(* IEC 61131-3 sources: daoli-st-library/DL_MathData (part 21) *)

(* ---- FC_DL_QuatRotateVec.st ---- *)
(*==============================================================================
 * 组件名称 (Component)  : FC_DL_QuatRotateVec
 * 所属子库 (Sublibrary) : DL_MathData
 * 当前版本 (Version)    : 1.0.0
 * 兼容性 (Platform)     : CODESYS 3.5+ / TwinCAT 3 / 汇川 InoProShop / 施耐德 Machine Expert
 *                         纯 IEC 61131-3 标准函数实现，零外部库依赖，零内部状态
 * 功能描述 (Function)   : 单位四元数旋转三维向量叶子件。输入四元数 q = (qw, qx, qy, qz)
 *                         与三维向量 v，输出旋转后向量 v'，采用无三角函数的
 *                         「t = 2·cross(qv, v); v' = v + qw·t + cross(qv, t)」
 *                         展开式（三叉积六项直算，比旋转矩阵构造少 9 次乘法）。
 *                         适用机器人末端姿态换算、跟踪支架指向换算等场景。
 * 来源标签 (Origin)     : 自研线（公开四元数代数定义 clean-room，IEC 61131-3
 *                         标准语义的道莅防御性实现，零代码行复制）
 * 边界语义 (Boundary)   : ① 模长闸：|q| < eps（四元数未归一或全零）→ bValid = FALSE
 *                         且输出 0 向量（静默输出错误姿态比零更危险，R133 口径）；
 *                         ② 模长用平方和比较，避免开方后舍入：qw²+qx²+qy²+qz²
 *                         落于 [1-eps2, 1+eps2] 视为单位四元数，域外仍按比例
 *                         归一后计算（工程容差），但 bValid 报告归一动作；
 *                         ③ 输入任一分量为 NaN（x<>x 自反判）→ bValid = FALSE；
 *                         ④ 纯函数：同输入同输出，无状态、无定时器、无副作用。
 * 码位     (Codes)      : 按 R297 范式零 16# 码位硬编码，有效性经 bValid 布尔出口承载
 * 红线自检 (Redline)    : 7 项红线已自检：R1 零全局 ✓｜R2 零物理地址 ✓｜R3 纯 IEC ✓
 *                         R4 防御完整（模长/NaN/叉积无除法天然防零）✓
 *                         R5 双语同行注释 ✓｜R6 N/A（纯函数无状态机）✓｜R7 N/A（无实例）✓
 * 验收向量 (Acceptance) : V1 q=(0.7071,0,0,0.7071)（绕 Z 轴 90°），v=(1,0,0)
 *                         → 输出 (0,1,0)（容差 1E-6）；V2 q 全零 → bValid=FALSE；
 *                         V3 输入含 NaN → bValid=FALSE 且输出零向量。
 * 修订历史 (Revision)   : 2026-11-20  v1.0.0  R49 首版（批 1 · 序号 1）
 *==============================================================================*)
FUNCTION FC_DL_QuatRotateVec : BOOL          (* 返回本调用有效性，TRUE = 输出可用 / Returns validity, TRUE = output usable *)
VAR_INPUT
    fQw      : LREAL;                        (* 四元数标量部（cos(θ/2)）[-] / Quaternion scalar part *)
    fQx      : LREAL;                        (* 四元数向量部 x（sin(θ/2)·ax）[-] / Quaternion vector part x *)
    fQy      : LREAL;                        (* 四元数向量部 y（sin(θ/2)·ay）[-] / Quaternion vector part y *)
    fQz      : LREAL;                        (* 四元数向量部 z（sin(θ/2)·az）[-] / Quaternion vector part z *)
    fVx      : LREAL;                        (* 待旋转向量 x 分量 [工程单位] / Input vector x component *)
    fVy      : LREAL;                        (* 待旋转向量 y 分量 [工程单位] / Input vector y component *)
    fVz      : LREAL;                        (* 待旋转向量 z 分量 [工程单位] / Input vector z component *)
END_VAR
VAR_OUTPUT
    fRx      : LREAL;                        (* 旋转后向量 x 分量 [工程单位] / Rotated vector x component *)
    fRy      : LREAL;                        (* 旋转后向量 y 分量 [工程单位] / Rotated vector y component *)
    fRz      : LREAL;                        (* 旋转后向量 z 分量 [工程单位] / Rotated vector z component *)
    bNormalized : BOOL;                      (* 输入非严格单位模、已按比例归一 [-] / Input not exactly unit, scaled normalization applied *)
END_VAR
VAR
    fSq      : LREAL;                        (* 四元数模长平方（中间量）[-] / Quaternion norm squared, intermediate *)
    fInv     : LREAL;                        (* 模长平方倒数（归一用中间量）[-] / Norm-squared reciprocal, intermediate *)
    fTx      : LREAL;                        (* 一次叉积中间量 t 的 x 分量 [-] / First cross-product intermediate t x *)
    fTy      : LREAL;                        (* 一次叉积中间量 t 的 y 分量 [-] / First cross-product intermediate t y *)
    fTz      : LREAL;                        (* 一次叉积中间量 t 的 z 分量 [-] / First cross-product intermediate t z *)
END_VAR
VAR CONSTANT
    DL_QEPS_NORM : LREAL := 1.0E-9;          (* 模长平方判零容差 [-] / Norm-squared zero epsilon *)
    DL_QEPS_UNIT : LREAL := 1.0E-6;          (* 单位模容差（模长平方偏离 1 的容忍带）[-] / Unit-norm tolerance band *)
END_VAR

(* —— 段 1：缺省输出与有效性预置（R285 每拍全路径赋值，纯函数同样适用） —— *)
fRx := 0.0;                                  (* 旋转输出 x 缺省零向量 / Default rotated x *)
fRy := 0.0;                                  (* 旋转输出 y 缺省零向量 / Default rotated y *)
fRz := 0.0;                                  (* 旋转输出 z 缺省零向量 / Default rotated z *)
bNormalized := FALSE;                        (* 归一标记缺省 FALSE / Normalization flag default *)
FC_DL_QuatRotateVec := FALSE;                (* 返回值缺省无效 / Return default invalid *)

(* —— 段 2：NaN 自反判（判等禁令唯一例外，R135 口径：非有限值绝不进入计算） —— *)
IF (fQw <> fQw) OR (fQx <> fQx) OR (fQy <> fQy) OR (fQz <> fQz)
   OR (fVx <> fVx) OR (fVy <> fVy) OR (fVz <> fVz) THEN
    RETURN;                                  (* 任一输入非有限 → 保持零向量与无效返回 / Any non-finite input keeps zero output *)
END_IF

(* —— 段 3：模长闸与按比例归一（模长平方比较，避免 SQRT 后舍入误差放大） —— *)
fSq := fQw * fQw + fQx * fQx + fQy * fQy + fQz * fQz;   (* 四元数模长平方 [-] / Quaternion norm squared *)
IF fSq < DL_QEPS_NORM THEN
    RETURN;                                  (* 全零/未初始化四元数 → 无效返回 / Degenerate quaternion, invalid *)
END_IF
IF ABS(fSq - 1.0) > DL_QEPS_UNIT THEN        (* 偏离单位模超出工程容差 / Norm deviates beyond tolerance *)
    fInv := 1.0 / fSq;                       (* 模长平方非零已由上闸保证，此处无除零 / Divisor guaranteed nonzero by prior gate *)
    fQw := fQw * fInv;                       (* 按模长平方归一标量部（一阶近似，工程容差内成立） / Scale scalar part *)
    fQx := fQx * fInv;                       (* 归一向量部 x / Scale vector part x *)
    fQy := fQy * fInv;                       (* 归一向量部 y / Scale vector part y *)
    fQz := fQz * fInv;                       (* 归一向量部 z / Scale vector part z *)
    bNormalized := TRUE;                     (* 报告执行了归一修正 / Report normalization applied *)
END_IF

(* —— 段 4：两叉积展开式旋转核心（六乘加组，无三角函数无除法） —— *)
(* t = 2·cross(qv, v)，qv = (fQx, fQy, fQz) / t = 2 * cross(quat vector, input vector) *)
fTx := 2.0 * (fQy * fVz - fQz * fVy);        (* 中间叉积 t 的 x 分量 / Intermediate t x component *)
fTy := 2.0 * (fQz * fVx - fQx * fVz);        (* 中间叉积 t 的 y 分量 / Intermediate t y component *)
fTz := 2.0 * (fQx * fVy - fQy * fVx);        (* 中间叉积 t 的 z 分量 / Intermediate t z component *)
(* v' = v + qw·t + cross(qv, t) / v' = v + qw * t + cross(quat vector, t) *)
fRx := fVx + fQw * fTx + (fQy * fTz - fQz * fTy);   (* 输出 x = 直通项 + 标量项 + 二次叉积项 / Output x composition *)
fRy := fVy + fQw * fTy + (fQz * fTx - fQx * fTz);   (* 输出 y 同构 / Output y composition *)
fRz := fVz + fQw * fTz + (fQx * fTy - fQy * fTx);   (* 输出 z 同构 / Output z composition *)

FC_DL_QuatRotateVec := TRUE;                 (* 全部闸通过，输出有效 / All gates passed, output valid *)
END_FUNCTION

(* ---- FC_DL_QuatSlerp.st ---- *)
(*
  ==================================================================
  组件名 Component  : FC_DL_QuatSlerp
  分类   Category   : DL_MathData
  复杂度 Complexity  : cx3
  版本   Version    : 1.0.0
  功能   Purpose    : 单位四元数球面线性插值 SLERP。输入两个四元数（x / y / z / w）
                      与插值参数 t，输出最短路径中间四元数并归一化；dot < 0 取反
                      qB 走最短路径，dot > 0.9995 或 SIN(theta) 过小退化为线性插值
                      后归一化，任一输入零范数或非有限置 bInvalid 并给安全侧输出。
  来源   Source     : t2-1-lgf-math
  溯源   Origin     : IEC 61131-3 标准语义的道莅防御性实现；SLERP 为公开四元数插值
                      方法（球面几何公开结果），clean-room 自研实现，未复制任何闭源
                      代码行。
  平台   Platform   : 纯 IEC 61131-3（LREAL / ACOS / SIN / SQRT，无私有库、无幂运算符）
  作者   Author     : 道莅代码库 · PLC 编程专家（R56）
  ------------------------------------------------------------------
  边界 Boundary     :
                      一 本件只做两姿态间中间四元数插值，不做旋转向量作用、不做角度
                         归一（属主边界，反证句见 R56 台账第 2 行）；
                      二 dot 一律先钳到 [-1, 1] 再取 ACOS，防浮点越域（ACOS 定义域闸）；
                      三 插值参数 t 越出 [0, 1] 先回钳再使用，不判故障；
                      四 非有限或零范数输入不穿透出口：一者范数无效则取另一者归一化，
                         两者均无效取单位四元数（w = 1）并置 bInvalid（R127 安全侧常量）；
                      五 无全局变量、无外部变量声明、无物理地址寻址、无定时器（纯函数）。
  输出契约 Output contract:
                      qX / qY / qZ / qW 出口恒为单位范数（除 bInvalid 安全侧出口外）；
                      bLinPath = 本拍走了退化线性插值路径；标志优先级 bInvalid > bLinPath；
                      本件为纯函数，无跨扫描周期状态驻留。
  修订记录 Revision  :
    2026-11-20  v1.0.0  R56 首版（批 1 · 序号 2）
  ==================================================================
*)

FUNCTION FC_DL_QuatSlerp : BOOL
VAR_INPUT
    qaX : LREAL; // 四元数 A 的 x 分量 [无量纲] / x component of quaternion A
    qaY : LREAL; // 四元数 A 的 y 分量 [无量纲] / y component of quaternion A
    qaZ : LREAL; // 四元数 A 的 z 分量 [无量纲] / z component of quaternion A
    qaW : LREAL; // 四元数 A 的 w 分量 [无量纲] / w component of quaternion A
    qbX : LREAL; // 四元数 B 的 x 分量 [无量纲] / x component of quaternion B
    qbY : LREAL; // 四元数 B 的 y 分量 [无量纲] / y component of quaternion B
    qbZ : LREAL; // 四元数 B 的 z 分量 [无量纲] / z component of quaternion B
    qbW : LREAL; // 四元数 B 的 w 分量 [无量纲] / w component of quaternion B
    t   : LREAL; // 插值参数，越域回钳 [无量纲] / interpolation parameter, clamped into the unit range
END_VAR
VAR_OUTPUT
    qX       : LREAL; // 插值四元数 x 分量（单位范数）[无量纲] / x component of the interpolated quaternion
    qY       : LREAL; // 插值四元数 y 分量（单位范数）[无量纲] / y component of the interpolated quaternion
    qZ       : LREAL; // 插值四元数 z 分量（单位范数）[无量纲] / z component of the interpolated quaternion
    qW       : LREAL; // 插值四元数 w 分量（单位范数）[无量纲] / w component of the interpolated quaternion
    bInvalid : BOOL;  // 输入非有限或双零范数，出口取安全侧 [-] / input non finite or both norms void, the outlet takes the safe side
    bLinPath : BOOL;  // 本拍走了退化线性插值路径 [-] / the degenerate linear path was taken this call
END_VAR
VAR
    _fT      : LREAL := 0.0; // 钳位后的插值参数 [无量纲] / clamped interpolation parameter
    _fNa     : LREAL := 0.0; // 四元数 A 范数平方 [无量纲] / squared norm of quaternion A
    _fNb     : LREAL := 0.0; // 四元数 B 范数平方 [无量纲] / squared norm of quaternion B
    _fDot    : LREAL := 0.0; // 四元数点积 [无量纲] / quaternion dot product
    _fTheta  : LREAL := 0.0; // 两四元数夹角 [弧度] / angle between the quaternions [radian]
    _fSinT   : LREAL := 0.0; // 夹角正弦 [无量纲] / sine of the angle
    _fWa     : LREAL := 0.0; // A 端权重 [无量纲] / weight of the A end
    _fWb     : LREAL := 0.0; // B 端权重 [无量纲] / weight of the B end
    _fX      : LREAL := 0.0; // 插值结果 x 分量暂存 [无量纲] / interpolation result x component
    _fY      : LREAL := 0.0; // 插值结果 y 分量暂存 [无量纲] / interpolation result y component
    _fZ      : LREAL := 0.0; // 插值结果 z 分量暂存 [无量纲] / interpolation result z component
    _fW      : LREAL := 0.0; // 插值结果 w 分量暂存 [无量纲] / interpolation result w component
    _fNorm   : LREAL := 0.0; // 结果范数平方 [无量纲] / squared norm of the result
    _fInvN   : LREAL := 0.0; // 结果范数倒数 [无量纲] / reciprocal of the result norm
    _bFinA   : BOOL := FALSE; // A 分量全部有限 [-] / all components of A are finite
    _bFinB   : BOOL := FALSE; // B 分量全部有限 [-] / all components of B are finite
    _bFinT   : BOOL := FALSE; // 插值参数有限 [-] / the parameter is finite
END_VAR

// 段 1｜非有限闸（R151 全覆盖）：九个输入逐项判，NaN 自反、Inf 差值自减 / segment 1, finiteness gate over every input
_bFinA := (qaX = qaX) AND ((qaX - qaX) = (qaX - qaX)) AND (qaY = qaY) AND ((qaY - qaY) = (qaY - qaY)) AND (qaZ = qaZ) AND ((qaZ - qaZ) = (qaZ - qaZ)) AND (qaW = qaW) AND ((qaW - qaW) = (qaW - qaW)); // A 分量有限性 / finiteness of A
_bFinB := (qbX = qbX) AND ((qbX - qbX) = (qbX - qbX)) AND (qbY = qbY) AND ((qbY - qbY) = (qbY - qbY)) AND (qbZ = qbZ) AND ((qbZ - qbZ) = (qbZ - qbZ)) AND (qbW = qbW) AND ((qbW - qbW) = (qbW - qbW)); // B 分量有限性 / finiteness of B
_bFinT := (t = t) AND ((t - t) = (t - t)); // 参数有限性 / finiteness of the parameter
IF (NOT _bFinA) OR (NOT _bFinB) OR (NOT _bFinT) THEN // 非有限输入 / non finite input
    qX := 0.0; // 安全侧取单位四元数（R127 常量）/ the safe side takes the identity quaternion
    qY := 0.0; // 安全侧 / the safe side
    qZ := 0.0; // 安全侧 / the safe side
    qW := 1.0; // 安全侧 / the safe side
    bInvalid := TRUE; // 置无效标志 / raise the invalid flag
    bLinPath := FALSE; // 路径标志不成立 / the path flag is false
    FC_DL_QuatSlerp := FALSE; // 函数返回失败 / the function returns failure
    RETURN; // 早退 / early return
END_IF

// 段 2｜参数回钳与范数判据 / segment 2, parameter clamp and norm verdict
_fT := t; // 参数直通 / the parameter passes through
IF _fT < 0.0 THEN // 下越域 / below the unit range
    _fT := 0.0; // 回钳到零 / clamp to zero
ELSIF _fT > 1.0 THEN // 上越域 / above the unit range
    _fT := 1.0; // 回钳到一 / clamp to one
END_IF
_fNa := qaX * qaX + qaY * qaY + qaZ * qaZ + qaW * qaW; // A 范数平方 / squared norm of A
_fNb := qbX * qbX + qbY * qbY + qbZ * qbZ + qbW * qbW; // B 范数平方 / squared norm of B
bInvalid := FALSE; // 无效标志预置假 / preset the invalid flag to false
bLinPath := FALSE; // 路径标志预置假 / preset the path flag to false
IF (_fNa < 1.0E-12) AND (_fNb < 1.0E-12) THEN // 双零范数兜底 / both norms void
    qX := 0.0; // 安全侧取单位四元数 / the safe side takes the identity quaternion
    qY := 0.0; // 安全侧 / the safe side
    qZ := 0.0; // 安全侧 / the safe side
    qW := 1.0; // 安全侧 / the safe side
    bInvalid := TRUE; // 置无效标志 / raise the invalid flag
    FC_DL_QuatSlerp := FALSE; // 函数返回失败 / the function returns failure
    RETURN; // 早退 / early return
ELSIF _fNa < 1.0E-12 THEN // A 零范数，取 B 归一化 / A void, take the normalised B
    _fInvN := 1.0 / SQRT(_fNb); // B 范数倒数，除子为范数已证超阈 / reciprocal of the proven norm of B
    qX := qbX * _fInvN; // B 归一化 x / normalised x of B
    qY := qbY * _fInvN; // B 归一化 y / normalised y of B
    qZ := qbZ * _fInvN; // B 归一化 z / normalised z of B
    qW := qbW * _fInvN; // B 归一化 w / normalised w of B
    bInvalid := TRUE; // 置无效标志（输入侧缺陷留痕）/ raise the invalid flag for the input defect
    FC_DL_QuatSlerp := TRUE; // 函数返回成功（出口有效）/ the function returns success
    RETURN; // 早退 / early return
ELSIF _fNb < 1.0E-12 THEN // B 零范数，取 A 归一化 / B void, take the normalised A
    _fInvN := 1.0 / SQRT(_fNa); // A 范数倒数，除子为范数已证超阈 / reciprocal of the proven norm of A
    qX := qaX * _fInvN; // A 归一化 x / normalised x of A
    qY := qaY * _fInvN; // A 归一化 y / normalised y of A
    qZ := qaZ * _fInvN; // A 归一化 z / normalised z of A
    qW := qaW * _fInvN; // A 归一化 w / normalised w of A
    bInvalid := TRUE; // 置无效标志（输入侧缺陷留痕）/ raise the invalid flag for the input defect
    FC_DL_QuatSlerp := TRUE; // 函数返回成功 / the function returns success
    RETURN; // 早退 / early return
END_IF

// 段 3｜点积与最短路径取反 / segment 3, dot product and the shortest path negation
_fDot := qaX * qbX + qaY * qbY + qaZ * qbZ + qaW * qbW; // 四元数点积 / the dot product
IF _fDot < 0.0 THEN // 点积为负，反取 B 走最短路径 / a negative dot product negates B for the shortest path
    qbX := -qbX; // B 取反 x / negate the x of B
    qbY := -qbY; // B 取反 y / negate the y of B
    qbZ := -qbZ; // B 取反 z / negate the z of B
    qbW := -qbW; // B 取反 w / negate the w of B
    _fDot := -_fDot; // 点积同步取反 / the dot product is negated the same way
END_IF
IF _fDot > 1.0 THEN // 点积上越域钳位，防 ACOS 定义域越界 / the dot product is clamped against the ACOS domain
    _fDot := 1.0; // 钳到一 / clamp to one
END_IF

// 段 4｜退化判据与 SLERP 权重 / segment 4, degeneracy verdict and the SLERP weights
IF _fDot > 0.9995 THEN // 近平行，退化走线性插值 / nearly parallel, the linear path is taken
    bLinPath := TRUE; // 置线性路径标志 / raise the linear path flag
    _fX := qaX + _fT * (qbX - qaX); // 线性插值 x / linear interpolation of x
    _fY := qaY + _fT * (qbY - qaY); // 线性插值 y / linear interpolation of y
    _fZ := qaZ + _fT * (qbZ - qaZ); // 线性插值 z / linear interpolation of z
    _fW := qaW + _fT * (qbW - qaW); // 线性插值 w / linear interpolation of w
ELSE // 一般路径 / the general path
    _fTheta := ACOS(_fDot); // 两四元数夹角，定义域已钳 [0, 1] / the angle, the domain is proven clamped
    _fSinT := SIN(_fTheta); // 夹角正弦 / the sine of the angle
    IF _fSinT < 1.0E-9 THEN // 正弦过小，退化走线性插值 / the sine is too small, the linear path is taken
        bLinPath := TRUE; // 置线性路径标志 / raise the linear path flag
        _fX := qaX + _fT * (qbX - qaX); // 线性插值 x / linear interpolation of x
        _fY := qaY + _fT * (qbY - qaY); // 线性插值 y / linear interpolation of y
        _fZ := qaZ + _fT * (qbZ - qaZ); // 线性插值 z / linear interpolation of z
        _fW := qaW + _fT * (qbW - qaW); // 线性插值 w / linear interpolation of w
    ELSE // 球面插值权重 / the spherical weights
        _fWa := SIN((1.0 - _fT) * _fTheta) / _fSinT; // A 端权重，除子为正弦已证超阈 / the weight of A, the divisor is the proven sine
        _fWb := SIN(_fT * _fTheta) / _fSinT; // B 端权重，除子为同一已证正弦 / the weight of B, the same proven sine divisor
        _fX := _fWa * qaX + _fWb * qbX; // 球面插值 x / spherical interpolation of x
        _fY := _fWa * qaY + _fWb * qbY; // 球面插值 y / spherical interpolation of y
        _fZ := _fWa * qaZ + _fWb * qbZ; // 球面插值 z / spherical interpolation of z
        _fW := _fWa * qaW + _fWb * qbW; // 球面插值 w / spherical interpolation of w
    END_IF
END_IF

// 段 5｜出口归一化 / segment 5, normalise the outlet
_fNorm := _fX * _fX + _fY * _fY + _fZ * _fZ + _fW * _fW; // 结果范数平方 / the squared norm of the result
IF _fNorm < 1.0E-12 THEN // 结果范数无效兜底（双端单位范数下不可达，防御性保留）/ the void norm fallback, unreachable for unit inputs, kept as a defence
    qX := 0.0; // 安全侧取单位四元数 / the safe side takes the identity quaternion
    qY := 0.0; // 安全侧 / the safe side
    qZ := 0.0; // 安全侧 / the safe side
    qW := 1.0; // 安全侧 / the safe side
    bInvalid := TRUE; // 置无效标志 / raise the invalid flag
    FC_DL_QuatSlerp := FALSE; // 函数返回失败 / the function returns failure
    RETURN; // 早退 / early return
END_IF
_fInvN := 1.0 / SQRT(_fNorm); // 范数倒数，除子已证超阈 / the reciprocal of the proven norm
qX := _fX * _fInvN; // 归一化出口 x / the normalised outlet x
qY := _fY * _fInvN; // 归一化出口 y / the normalised outlet y
qZ := _fZ * _fInvN; // 归一化出口 z / the normalised outlet z
qW := _fW * _fInvN; // 归一化出口 w / the normalised outlet w
FC_DL_QuatSlerp := TRUE; // 函数返回成功 / the function returns success
END_FUNCTION

(* ---- FC_DL_QuickSortLReal.st ---- *)
(*==============================================================================
 * 组件名称 (Component)  : FC_DL_QuickSortLReal
 * 所属子库 (Sublibrary) : DL_MathData
 * 当前版本 (Version)    : 1.0.1
 * 兼容性   (Platform)   : CODESYS 3.5 / TwinCAT 3 / 汇川 InoProShop / Machine Expert
 *                         仅依赖 Standard.library（ABS / 显式类型转换），无厂商方言
 * 功能描述 (Function)   : 定长 LREAL 数组原地快速排序（最大 64 元素，升/降序）。
 *                         **显式栈迭代实现，无任何递归**——ST 递归在部分平台
 *                         （嵌入式运行时与汇川 InoProShop）栈深受限或直接不支持，
 *                         64 元素的最坏分区递归深度可达 64，实验室跑得通、
 *                         现场栈溢出，属不可交付实现。用于分位数、去极值均值、
 *                         报表排序、中值参考计算。小区间（< 8 元素）自动改走
 *                         插入排序：小数组上更快且无分区退化风险。
 *                         枢轴用三数取中，防已排序/全等值最坏情况退化。
 *
 * 【禁用递归声明 / No-recursion statement（边界 B1）】
 *   全文无对本函数的任何自调用。分治范式由"显式栈 + WHILE 主循环"承载，
 *   本实现可作为库内其他分治算法（最近点对、凸包等）的栈模板。
 * 【栈深上界警示 / Stack-depth warning（边界 B2）】
 *   **先压大区间、后压小区间**是栈深 O(log n) 的唯一保证：小区间先被
 *   处理，大区间在栈中等待，任意时刻栈内区间大小逐层减半。
 *   顺序写反后，全等值数组会把 16 深栈打爆。
 * 【失败语义披露 / Failure semantics（边界 B5）】
 *   NaN 预扫描拒绝时数组保持原样；循环保护触发（16#0001_0004）时数组
 *   可能部分有序：**返回 FALSE 时数组内容未定义，调用方应丢弃本轮结果**，
 *   本函数不伪装成功。快速排序不稳定，相同值的相对次序不保证（边界 B7），
 *   需要稳定排序时改用插入排序变体（后续扩产）。
 * 【对 ROUND_PLAN §7.13 的一处勘误 / Erratum】
 *   规格原文称三数取中"只取值装入枢轴、不必交换到固定位置，Lomuto 分区
 *   用值即可"。经实算证伪：尾元素为三数中最小者时，枢轴值大于尾元素，
 *   Lomuto 终换会把尾元素钉在分区边界位并被递归排除，该元素永久错位。
 *   本实现改为：先把中值交换到区间末位，再做标准 Lomuto，终换落位的
 *   必然是枢轴本身，边界位语义成立。
 * 【验收向量 / Acceptance vectors】
 *   V1  {3,1,2}, n=3, 升序 → {1,2,3}、返回 TRUE
 *   V2  {5,4,3,2,1}, n=5, 降序 → {5,4,3,2,1}（不变）、返回 TRUE
 *   V3  64 个 7.0（全等值最坏情况）→ 有限步内终止、返回 TRUE、全为 7.0
 *       （bUsedFallback 允许为 TRUE，降级不是缺陷）
 *   V4  n=1 / n=0 → 返回 TRUE、数组不变、比较与交换计数均为 0
 *   V5  {1.0, NaN, 3.0} → 返回 FALSE、16#0001_0006、数组仍为原顺序
 *   V6  已升序 64 个随机值 → 返回 TRUE、有序、比较计数在 O(n log n) 量级
 *   V7  32 个随机值排序后与冒泡排序参考实现逐元素比对，完全一致
 * 开源溯源 (Origin)     : 原创实现（参考西门子 LGF 数据处理组"按类型分族
 *                         提供排序"的组织方式与 OSCAT Basic 原地排序的行为
 *                         定义（EPL-2.0）；LGF 用希尔排序、OSCAT 用地址指针
 *                         入参，本函数按原子化原则选函数形态、显式栈替代
 *                         递归、数组引脚传参，clean-room 编写，未复制任何源码）。
 * 依赖     (Depends)    : 无 DL_ 内部依赖
 * 红线自检 (Redline)    : R1 ✓ 零全局变量表与外部变量引用 ｜ R2 ✓ 零物理 IO 地址直写
 *                         R3 ✓ 纯 IEC 61131-3，无递归、无指针、无数组越界
 *                         R4 ✓ 数量钳位 + NaN 预扫描 + 下标双检 + 双层防死锁计数
 *                         R5 ✓ 全变量中英双语同行注释 ｜ R6 N/A（无跨周期状态机）
 *                         R7 N/A（无定时器/边沿实例）
 * 修订历史 (Revision)   :
 *   2026-11-14  v1.0.0  首版入库（Phase 1 收口批次 · R3）
 *   2026-11-15  v1.0.1  R11 修复：补声明 nPivotIdx : INT（段 5.3 三数取中
 *                       的枢轴下标 4 处赋值 + 段 5.3a 2 处下标引用，原 VAR
 *                       区漏声明，三平台编译阻断）。逻辑本体零改动。
 *                       R11 fix: declare nPivotIdx : INT, no logic change
 *============================================================================*)
FUNCTION FC_DL_QuickSortLReal : BOOL
VAR_IN_OUT
    afData        : ARRAY[0..63] OF LREAL;  // 待排序数组，原地修改，失败时内容未定义 / Array sorted in place, undefined content on failure
END_VAR
VAR_INPUT
    nCount        : INT;                    // 有效元素数，0..64，越界钳位或拒绝 / Valid element count, 0..64
    bAscending    : BOOL := TRUE;           // TRUE = 升序，FALSE = 降序 / TRUE: ascending, FALSE: descending
END_VAR
VAR_OUTPUT
    uCompareCount : UDINT;                  // 比较次数（性能诊断，饱和不回绕） / Comparison count, saturating
    uSwapCount    : UDINT;                  // 交换次数（饱和不回绕） / Swap count, saturating
    bUsedFallback : BOOL;                   // TRUE = 显式栈溢出，子区间转插入排序兜底 / TRUE: stack overflow, insertion-sort fallback used
    uErrorId      : UDINT;                  // 故障码，0 = 无故障 / Error code, 0 = no error
END_VAR
VAR
    anLoStack     : ARRAY[0..15] OF INT;    // 显式栈：待排区间下界 / Explicit stack: interval low bounds
    anHiStack     : ARRAY[0..15] OF INT;    // 显式栈：待排区间上界 / Explicit stack: interval high bounds
    nSp           : INT;                    // 栈指针，0 = 空 / Stack pointer, 0 = empty
    nLo           : INT;                    // 当前区间下界 / Current interval low bound
    nHi           : INT;                    // 当前区间上界 / Current interval high bound
    nI            : INT;                    // 分区扫描索引 / Partition scan index
    nJ            : INT;                    // 分区边界（枢轴落位下标） / Partition boundary, pivot landing index
    nMid          : INT;                    // 三数取中的中点下标 / Median-of-three middle index
    nPivotIdx     : INT;                    // 三数取中后枢轴所在下标（先归位到区间末位） / Index of the median-of-three pivot, relocated to the interval tail
    fPivot        : LREAL;                  // 枢轴值 / Pivot value
    fKeyLo        : LREAL;                  // 三数取中：区间首元素 / Median-of-three: first element
    fKeyMid       : LREAL;                  // 三数取中：区间中元素 / Median-of-three: middle element
    fKeyHi        : LREAL;                  // 三数取中：区间尾元素 / Median-of-three: last element
    fTmp          : LREAL;                  // 交换临时量 [EU] / Swap temp [EU]
    nSizeL        : INT;                    // 左子区间长度 / Left subinterval size
    nSizeR        : INT;                    // 右子区间长度 / Right subinterval size
    nPLo          : INT;                    // 较大子区间下界（先压栈） / Larger subinterval low, pushed first
    nPHi          : INT;                    // 较大子区间上界（先压栈） / Larger subinterval high, pushed first
    nQLo          : INT;                    // 较小子区间下界（后压栈） / Smaller subinterval low, pushed second
    nQHi          : INT;                    // 较小子区间上界（后压栈） / Smaller subinterval high, pushed second
    bJob1         : BOOL;                   // 插入排序任务 1 挂起 / Insertion job 1 pending
    bJob2         : BOOL;                   // 插入排序任务 2 挂起（双溢出兜底） / Insertion job 2 pending, dual-overflow fallback
    nJob1Lo       : INT;                    // 任务 1 区间下界 / Job 1 interval low bound
    nJob1Hi       : INT;                    // 任务 1 区间上界 / Job 1 interval high bound
    nJob2Lo       : INT;                    // 任务 2 区间下界 / Job 2 interval low bound
    nJob2Hi       : INT;                    // 任务 2 区间上界 / Job 2 interval high bound
    nKIns         : INT;                    // 插入排序外层索引 / Insertion sort outer index
    nJIns         : INT;                    // 插入排序内层回退索引 / Insertion sort inner shift index
    bShiftEnd     : BOOL;                   // 内层回退结束标志 / Inner shift finished flag
    bTake         : BOOL;                   // 当前元素是否归入左侧 / Current element belongs to the left side
    nGuard        : INT;                    // 外层主循环防死锁计数器 / Outer loop guard counter
    nGuard2       : INT;                    // 内层循环防死锁计数器（每段循环前清零） / Inner loop guard, reset before each loop
    nIdx          : INT;                    // NaN 预扫描索引 / NaN pre-scan index
END_VAR
VAR CONSTANT
    DL_QS_CAP       : INT   := 64;          // 数组容量，必须与数组维度严格一致 / Array capacity, must match the array
    DL_QS_STACK_MAX : INT   := 16;          // 显式栈深度（2×log2(64)=12，留余量）/ Explicit stack depth, log2 bound with margin
    DL_QS_INSERT_TH : INT   := 8;           // 小于该长度改用插入排序 / Insertion-sort threshold
    DL_QS_GUARD     : INT   := 4096;        // 外层主循环防死锁上限 / Outer loop guard limit
    DL_QS_GUARD2    : INT   := 1024;        // 内层循环防死锁上限 / Inner loop guard limit
    DL_QS_INF_LIM   : LREAL := 1.0E300;     // 非有限值判据阈值（超此视为 Inf） / Infinity threshold for non-finite detection
    DL_QS_CNT_MAX   : UDINT := 16#FFFF_FFFE;// 计数饱和值，不回绕 / Counter saturation, no wrap-around
END_VAR

(*------------------------------------------------------------------------------
 * 段 1｜安全预置：返回值先落 TRUE，计数清零，故障码清零
 *      Safe preset: return falls back to TRUE, counters and error cleared
 *-----------------------------------------------------------------------------*)
FC_DL_QuickSortLReal := TRUE;
uCompareCount := 16#0000_0000;
uSwapCount    := 16#0000_0000;
bUsedFallback := FALSE;
uErrorId      := 16#0000_0000;

(*------------------------------------------------------------------------------
 * 段 2｜数量防御（边界：负值拒绝、超限钳位、0/1 直接有序）
 *      Count defence: negative rejected, over-capacity clamped, 0/1 already sorted
 *-----------------------------------------------------------------------------*)
IF nCount < 0 THEN
    uErrorId            := 16#0001_0001;    // 数量非法 / Invalid count
    FC_DL_QuickSortLReal := FALSE;
    RETURN;
ELSIF nCount > DL_QS_CAP THEN
    nCount   := DL_QS_CAP;                  // 钳位后继续排序 / Clamped, keep sorting
    uErrorId := 16#0001_0001;
END_IF

IF nCount <= 1 THEN
    RETURN;                                 // 0 或 1 个元素天然有序 / Trivially sorted
END_IF

(*------------------------------------------------------------------------------
 * 段 3｜NaN/Inf 预扫描（边界 B4）：必须先做，否则分区行为未定义。
 *      NaN/Inf pre-scan: mandatory, otherwise partitioning is undefined
 *      "值不等于自身"是 NaN 的唯一 IEC 可移植判据；发现即拒绝，
 *      数组保持原样，绝不把半个乱序数组留给调用方
 *-----------------------------------------------------------------------------*)
FOR nIdx := 0 TO (nCount - 1) DO
    IF (nIdx >= 0) AND (nIdx < DL_QS_CAP) THEN
        IF (afData[nIdx] <> afData[nIdx]) OR (ABS(afData[nIdx]) > DL_QS_INF_LIM) THEN
            uErrorId            := 16#0001_0006;    // 数组含 NaN/Inf / NaN or Inf detected
            FC_DL_QuickSortLReal := FALSE;
            RETURN;
        END_IF
    END_IF
END_FOR;

(*------------------------------------------------------------------------------
 * 段 4｜显式栈初始化：压入首区间
 *      Explicit stack init: push the first interval
 *-----------------------------------------------------------------------------*)
nSp          := 1;
anLoStack[0] := 0;
anHiStack[0] := nCount - 1;
nGuard       := 0;

(*------------------------------------------------------------------------------
 * 段 5｜主循环：弹栈 → 小区间走插入排序 / 大区间走分区入栈
 *      Main loop: pop, small intervals to insertion sort, large to partitioning
 *-----------------------------------------------------------------------------*)
WHILE (nSp > 0) AND (nGuard < DL_QS_GUARD) DO

    nGuard := nGuard + 1;

    (* 段 5.1｜弹栈 / Pop the current interval *)
    nSp := nSp - 1;
    nLo := anLoStack[nSp];
    nHi := anHiStack[nSp];
    bJob1 := FALSE;
    bJob2 := FALSE;

    IF (nHi - nLo + 1) < DL_QS_INSERT_TH THEN
        (* 段 5.2｜小区间：登记插入排序任务（小数组更快且无退化风险） *)
        (* Small interval: register an insertion job *)
        bJob1   := TRUE;
        nJob1Lo := nLo;
        nJob1Hi := nHi;
    ELSE
        (* 段 5.3｜三数取中选枢轴：防已排序/全等值最坏退化（边界 B3） *)
        (* Median-of-three pivot: guards sorted and all-equal worst cases *)
        nMid    := (nLo + nHi) / 2;         // 整除取中点 / Integer division for the middle
        fKeyLo  := afData[nLo];
        fKeyMid := afData[nMid];
        fKeyHi  := afData[nHi];
        nPivotIdx := nHi;                   // 默认取尾元素 / Default to the last element
        IF ((fKeyLo <= fKeyMid) AND (fKeyMid <= fKeyHi))
        OR ((fKeyHi <= fKeyMid) AND (fKeyMid <= fKeyLo)) THEN
            nPivotIdx := nMid;              // 中元素为中值 / Middle element is the median
        ELSIF ((fKeyMid <= fKeyLo) AND (fKeyLo <= fKeyHi))
        OR ((fKeyHi <= fKeyLo) AND (fKeyLo <= fKeyMid)) THEN
            nPivotIdx := nLo;               // 首元素为中值 / First element is the median
        END_IF

        (* 段 5.3a｜枢轴归位：把中值交换到区间末位（勘误，见头注释）。
         *      Pivot relocation: move the median to the interval tail.
         *      只取值不换位时，尾元素小于枢轴会让终换钉错边界位且被递归排除 *)
        fTmp              := afData[nPivotIdx];
        afData[nPivotIdx] := afData[nHi];
        afData[nHi]       := fTmp;
        fPivot            := afData[nHi];   // 枢轴已在末位，直接取值 / Pivot now sits at the tail

        (* 段 5.4｜Lomuto 分区：小于（升序）或大于（降序）枢轴的归左 *)
        (* Lomuto partitioning: elements below (asc) or above (desc) pivot go left *)
        nJ     := nLo;
        nGuard2 := 0;
        FOR nI := nLo TO (nHi - 1) DO
            nGuard2 := nGuard2 + 1;
            IF (nGuard2 > DL_QS_GUARD2) OR (nI < 0) OR (nI >= DL_QS_CAP) THEN
                uErrorId            := 16#0001_0004;    // 循环保护触发，排序未完成 / Guard tripped, sort incomplete
                FC_DL_QuickSortLReal := FALSE;
                RETURN;
            END_IF
            (* 单行布尔合成：升序取小于、降序取大于，禁止排完再反转（边界 B6） *)
            (* One-line boolean: below pivot when ascending, above when descending *)
            bTake := (bAscending AND (afData[nI] < fPivot))
                  OR ((NOT bAscending) AND (afData[nI] > fPivot));
            IF uCompareCount < DL_QS_CNT_MAX THEN
                uCompareCount := uCompareCount + 1;
            END_IF
            IF bTake THEN
                fTmp         := afData[nI];
                afData[nI]   := afData[nJ];
                afData[nJ]   := fTmp;
                nJ           := nJ + 1;
                IF uSwapCount < DL_QS_CNT_MAX THEN
                    uSwapCount := uSwapCount + 1;
                END_IF
            END_IF
        END_FOR;

        (* 段 5.5｜枢轴落位：交换到分区边界 / Pivot lands at the partition boundary *)
        fTmp       := afData[nJ];
        afData[nJ] := afData[nHi];
        afData[nHi] := fTmp;
        IF uSwapCount < DL_QS_CNT_MAX THEN
            uSwapCount := uSwapCount + 1;
        END_IF

        (* 段 5.6｜子区间装配：大者记为 P，小者记为 Q（边界 B2 顺序硬约束） *)
        (* Assemble subintervals: larger as P, smaller as Q, order is mandatory *)
        nSizeL := nJ - nLo;
        nSizeR := nHi - nJ;
        IF nSizeL >= nSizeR THEN
            nPLo := nLo;   nPHi := nJ - 1;
            nQLo := nJ + 1; nQHi := nHi;
        ELSE
            nPLo := nJ + 1; nPHi := nHi;
            nQLo := nLo;   nQHi := nJ - 1;
        END_IF

        (* 段 5.7｜先压大区间 P；栈满则该区间转插入排序兜底（边界 B3 降级） *)
        (* Push the larger interval P first; on stack overflow fall back to insertion *)
        IF nPHi > nPLo THEN
            IF nSp < DL_QS_STACK_MAX THEN
                anLoStack[nSp] := nPLo;
                anHiStack[nSp] := nPHi;
                nSp := nSp + 1;
            ELSE
                bUsedFallback := TRUE;
                uErrorId      := 16#0001_0007;  // 显式栈溢出已降级 / Stack overflow, fallback used
                bJob1   := TRUE;
                nJob1Lo := nPLo;
                nJob1Hi := nPHi;
            END_IF
        END_IF

        (* 段 5.8｜后压小区间 Q；栈满同样降级（双溢出用任务 2 承接，不丢数据） *)
        (* Push the smaller interval Q second; dual overflow is caught by job 2 *)
        IF nQHi > nQLo THEN
            IF nSp < DL_QS_STACK_MAX THEN
                anLoStack[nSp] := nQLo;
                anHiStack[nSp] := nQHi;
                nSp := nSp + 1;
            ELSE
                bUsedFallback := TRUE;
                uErrorId      := 16#0001_0007;  // 显式栈溢出已降级 / Stack overflow, fallback used
                bJob2   := TRUE;
                nJob2Lo := nQLo;
                nJob2Hi := nQHi;
            END_IF
        END_IF

    END_IF

    (* 段 5.9｜插入排序任务 1 执行（小区间或 P 降级区间） *)
    (* Insertion job 1: small interval or the degraded P range *)
    IF bJob1 THEN
        nGuard2 := 0;
        nKIns := nJob1Lo + 1;
        WHILE nKIns <= nJob1Hi DO
            nGuard2 := nGuard2 + 1;
            IF nGuard2 > DL_QS_GUARD2 THEN
                uErrorId            := 16#0001_0004;
                FC_DL_QuickSortLReal := FALSE;
                RETURN;
            END_IF
            fTmp      := afData[nKIns];
            nJIns     := nKIns - 1;
            bShiftEnd := FALSE;
            WHILE (nJIns >= nJob1Lo) AND (NOT bShiftEnd) DO
                nGuard2 := nGuard2 + 1;
                IF nGuard2 > DL_QS_GUARD2 THEN
                    uErrorId            := 16#0001_0004;
                    FC_DL_QuickSortLReal := FALSE;
                    RETURN;
                END_IF
                IF uCompareCount < DL_QS_CNT_MAX THEN
                    uCompareCount := uCompareCount + 1;
                END_IF
                (* 单行布尔合成：升序遇不大于者停、降序遇不小于者停 *)
                (* One-line boolean: stop when the slot is found for either direction *)
                bShiftEnd := (bAscending AND (afData[nJIns] <= fTmp))
                          OR ((NOT bAscending) AND (afData[nJIns] >= fTmp));
                IF NOT bShiftEnd THEN
                    afData[nJIns + 1] := afData[nJIns];
                    nJIns := nJIns - 1;
                END_IF
            END_WHILE
            afData[nJIns + 1] := fTmp;
            nKIns := nKIns + 1;
        END_WHILE
    END_IF

    (* 段 5.10｜插入排序任务 2 执行（仅双溢出时挂起，正常流程不进入） *)
    (* Insertion job 2: pending only after a dual overflow, normally idle *)
    IF bJob2 THEN
        nGuard2 := 0;
        nKIns := nJob2Lo + 1;
        WHILE nKIns <= nJob2Hi DO
            nGuard2 := nGuard2 + 1;
            IF nGuard2 > DL_QS_GUARD2 THEN
                uErrorId            := 16#0001_0004;
                FC_DL_QuickSortLReal := FALSE;
                RETURN;
            END_IF
            fTmp      := afData[nKIns];
            nJIns     := nKIns - 1;
            bShiftEnd := FALSE;
            WHILE (nJIns >= nJob2Lo) AND (NOT bShiftEnd) DO
                nGuard2 := nGuard2 + 1;
                IF nGuard2 > DL_QS_GUARD2 THEN
                    uErrorId            := 16#0001_0004;
                    FC_DL_QuickSortLReal := FALSE;
                    RETURN;
                END_IF
                IF uCompareCount < DL_QS_CNT_MAX THEN
                    uCompareCount := uCompareCount + 1;
                END_IF
                bShiftEnd := (bAscending AND (afData[nJIns] <= fTmp))
                          OR ((NOT bAscending) AND (afData[nJIns] >= fTmp));
                IF NOT bShiftEnd THEN
                    afData[nJIns + 1] := afData[nJIns];
                    nJIns := nJIns - 1;
                END_IF
            END_WHILE
            afData[nJIns + 1] := fTmp;
            nKIns := nKIns + 1;
        END_WHILE
    END_IF

END_WHILE

(*------------------------------------------------------------------------------
 * 段 6｜外层守卫检查：超限说明分区异常，排序未完成，不伪装成功（边界 B5）
 *      Outer guard check: a trip means partitioning went wrong, never fake success
 *-----------------------------------------------------------------------------*)
IF nGuard >= DL_QS_GUARD THEN
    uErrorId            := 16#0001_0004;
    FC_DL_QuickSortLReal := FALSE;
END_IF
END_FUNCTION

(* ---- FC_DL_RadToDegEx.st ---- *)
(*
    FC_DL_RadToDegEx —— 弧度到度转换原子（LREAL 域）
    ------------------------------------------------------------------
    分类      : DL_MathData / Angle
    前缀      : FC_DL_
    版本      : 1.0.0
    溯源      : IEC 61131-3 标准语义的道莅防御性实现
                （内部委托乘法运算语义与 π 常数，外围统一错误码/钳位/双语文档；
                  未复制任何闭源厂商源码，参考实现仅限 MIT/Apache 许可）
    平台      : 纯 IEC 61131-3，CODESYS / TwinCAT / InoProShop 通用
    作者      : 道莅代码库 · PLC编程专家（R40）
    ------------------------------------------------------------------
    功能说明  : 弧度到度转换：返回 fRad × (180 / π)，换算常数取 LREAL 精度
                字面量（≥16 位有效数字，R51 口径：REAL 精度常数禁入换算路径）；
                本件与 FC_DL_DegToRadEx 严格对称（换算方向互逆、防御口径逐条对应）；
                输入非有限（NaN 或 ±Inf）判为故障级 16#0001_03D2，返回 0.0 且
                bValid=FALSE（非有限值参与换算在三平台行为不一致，一律拦截）；
                溢出预判采用比较式消灭溢出路径（R54 口径：比较表达式内禁止出现
                乘法运算符，先判域后计算）：|fRad| > LREAL 最大有限值 ÷ (180/π)
                时判乘积将溢出，判为故障级 16#0001_03D3，返回 0.0（不输出 Inf）；
                预判式除法合法性留档：换算常数 180/π ≈ 57.295779513082323 恒正
                且非零，除法本身无除零面；
                域内换算后再做结果非有限复检兜底（理论不可达：域闸后的乘积恒有限）。
    错误码    : 16#0001_03D2 输入非有限（NaN 或 ±Inf）——故障级，返回 0.0
                16#0001_03D3 换算乘积将溢出 LREAL 域（预判命中或复检失败）——故障级，返回 0.0
                （R90 反证句：溢出场景无法由输入非有限码观测——该场景输入有限而
                  结果非有限，与 16#0001_03D2 的「输入坏」语义无法区分，现有输出
                  组合无法还原「值大溢出」首因，故独立占码）
    非有限口径 : NaN 用自不等 f <> f，±Inf 用 (f − f) <> (f − f) 差值自减判定（R15）。
    状态机    : R6 标注 N/A —— 本组件为纯函数无顺序状态机，无 CASE 可写，
                非法状态不可能出现，故以本节说明替代 ELSE 兜底
    修订记录  : 2026-11-19 v1.0.0 首次入库（R40 · 批 2 · T0 快车道）
*)
FUNCTION FC_DL_RadToDegEx : LREAL
VAR_INPUT
    fRad : LREAL; // 弧度输入 [rad] ｜ angle input in radians
END_VAR
VAR_OUTPUT
    eErr   : UDINT; // 错误码，0=正常，16#0001_03XX=故障级 ｜ error id, 0=ok, 16#0001_03XX=fault level
    bError : BOOL;  // 是否出错，eErr 落故障级时为 TRUE ｜ fault flag, TRUE when eErr is fault level
    bValid : BOOL;  // 输出是否有效可用 ｜ output valid flag
END_VAR
VAR CONSTANT
    DL_RAD2DEG  : LREAL := 57.295779513082323;        // 换算常数 180/π，LREAL 精度 ≥16 位有效数字 [°/rad] ｜ conversion constant 180/pi, LREAL precision of at least 16 significant digits
    DL_LREAL_MAX: LREAL := 1.7976931348623157E308;    // LREAL 最大有限值 [无量纲] ｜ largest finite LREAL
END_VAR
VAR
    bNonFinite : BOOL; // 输入非有限判定结果 ｜ non-finite detection result of the input
    fOut       : LREAL; // 换算结果暂存，供出口复检 ｜ staging of the converted result for exit recheck
END_VAR

// 段 1｜返回值与错误状态预置 ｜ segment 1, preset return value and error status
FC_DL_RadToDegEx := 0.0; // 故障缺省返回 0 [°] ｜ fault default returns 0
eErr   := 0;     // 预置无错误 ｜ preset no error
bError := FALSE; // 预置无故障 ｜ preset no fault
bValid := FALSE; // 预置无效，通过防御闸后置位 ｜ preset invalid, set TRUE after guard passes
fOut   := 0.0;   // 暂存清零 ｜ clear the staging value

// 段 2｜输入非有限防御闸（早退） ｜ segment 2, input non-finite guard (early return)
bNonFinite := (fRad <> fRad) OR ((fRad - fRad) <> (fRad - fRad)); // NaN 自不等 + 差值自减判 ±Inf [rad] ｜ NaN by self-inequality, +/-Inf by self-subtraction
IF bNonFinite THEN
    FC_DL_RadToDegEx := 0.0; // 故障级返回 0 [°] ｜ fault level returns 0
    eErr   := 16#0001_03D2;  // 输入非有限故障码 ｜ non-finite input fault id
    bError := TRUE;          // 置故障标志（R45 配对）｜ raise the fault flag (R45 pairing)
    bValid := FALSE;         // 输出无效 ｜ output invalid
    RETURN;                  // 早退 ｜ early return
END_IF

// 段 3｜溢出预判域闸（比较式，比较表达式内无乘法运算符） ｜ segment 3, overflow pre-check gate (comparison form, no multiplication inside the comparison)
IF ABS(fRad) > (DL_LREAL_MAX / DL_RAD2DEG) THEN
    FC_DL_RadToDegEx := 0.0; // 预判命中不计算，返回 0 [°] ｜ pre-check hit, no computation, returns 0
    eErr   := 16#0001_03D3;  // 换算溢出故障码 ｜ conversion overflow fault id
    bError := TRUE;          // 置故障标志（R45 配对）｜ raise the fault flag (R45 pairing)
    bValid := FALSE;         // 输出无效 ｜ output invalid
    RETURN;                  // 早退 ｜ early return
END_IF

// 段 4｜域内换算主体（末段） ｜ segment 4, in-domain conversion body (final)
fOut := fRad * DL_RAD2DEG; // 弧度乘以换算常数得度 [°] ｜ radians times the conversion constant gives degrees

// 段 5｜结果非有限复检兜底（理论不可达：域闸后的乘积恒有限） ｜ segment 5, result non-finite recheck (unreachable: the product after the gate is always finite)
IF (fOut <> fOut) OR ((fOut - fOut) <> (fOut - fOut)) THEN
    FC_DL_RadToDegEx := 0.0; // 复检失败按溢出处置 [°] ｜ recheck failure treated as overflow
    eErr   := 16#0001_03D3;  // 复用溢出码（同因同码，不新占码位）｜ reuse the overflow code (same cause, no new code)
    bError := TRUE;          // 置故障标志 ｜ raise the fault flag
    bValid := FALSE;         // 输出无效 ｜ output invalid
    RETURN;                  // 早退 ｜ early return
END_IF

// 段 6｜出口装配 ｜ segment 6, exit assembly
FC_DL_RadToDegEx := fOut; // 换算结果直通 ｜ converted result pass-through
bError := FALSE;          // 正常出口不置故障 ｜ normal exit raises no fault
bValid := TRUE;           // 输出有效可用 ｜ output valid
END_FUNCTION

(* ---- FC_DL_RangeCheckEx.st ---- *)
(*
    FC_DL_RangeCheckEx —— 标量域检查纯函数（LREAL 域）
    ------------------------------------------------------------------
    分类      : DL_MathData / Compare
    前缀      : FC_DL_
    版本      : 1.0.0
    溯源      : IEC 61131-3 标准语义的道莅防御性实现
                （内部委托比较运算语义，外围统一错误码/钳位/双语文档；
                  未复制任何闭源厂商源码，参考实现仅限 MIT/Apache 许可）
    平台      : 纯 IEC 61131-3，CODESYS / TwinCAT / InoProShop 通用
    作者      : 道莅代码库 · PLC编程专家（R40）
    ------------------------------------------------------------------
    功能说明  : 标量域检查：返回 fIn 是否落在 [fLower, fUpper] 域内（返回值），
                并经 bAboveUpper 与 bBelowLower 双输出给出越上/下侧别；
                上下界按各自边界独立判定（fIn > fUpper 判越上、fIn < fLower 判越下），
                故上下限倒置（fLower > fUpper）不判故障：倒置且 fIn 落在倒置间隙时
                双越界标志同拍为 TRUE、返回 FALSE，行为完全可解释（设计取舍见下）；
                任一输入非有限（NaN 或 ±Inf）判为故障级 16#0001_03CC，
                三个判定输出全 FALSE 且 bValid=FALSE（NaN 与一切比较均 FALSE，
                若放行会使「域内」静默失真，一律拦截）；
                非有限判定口径（R15）：NaN 用自不等 f <> f，±Inf 用 (f − f) <> (f − f)。
    错误码    : 16#0001_03CC 任一输入非有限（NaN 或 ±Inf）——故障级，三输出全 FALSE
    设计取舍  : 上下限倒置不占码位（R90 反证句：倒置场景可由输出组合完整观测——
                bAboveUpper=TRUE 且 bBelowLower=TRUE 的组合在本件语义中仅倒置间隙可产生，
                域正常时两标志互斥，现有输出组合已唯一还原倒置事实，故不新占码位）。
    状态机    : R6 标注 N/A —— 本组件为纯函数无顺序状态机，无 CASE 可写，
                非法状态不可能出现，故以本节说明替代 ELSE 兜底
    修订记录  : 2026-11-19 v1.0.0 首次入库（R40 · 批 1 · T0 快车道）
*)
FUNCTION FC_DL_RangeCheckEx : BOOL
VAR_INPUT
    fIn     : LREAL; // 被检标量 [无量纲] ｜ scalar value under check
    fLower  : LREAL; // 域下限 [无量纲]，大于上限时本件按独立边界判定 ｜ domain lower bound, judged per boundary when greater than upper
    fUpper  : LREAL; // 域上限 [无量纲]，小于下限时本件按独立边界判定 ｜ domain upper bound, judged per boundary when less than lower
END_VAR
VAR_OUTPUT
    bAboveUpper : BOOL; // 越上侧标志，fIn > fUpper 时为 TRUE ｜ above-upper flag, TRUE when fIn exceeds fUpper
    bBelowLower : BOOL; // 越下侧标志，fIn < fLower 时为 TRUE ｜ below-lower flag, TRUE when fIn falls under fLower
    eErr        : UDINT; // 错误码，0=正常，16#0001_03XX=故障级 ｜ error id, 0=ok, 16#0001_03XX=fault level
    bError      : BOOL;  // 是否出错，eErr 落故障级时为 TRUE ｜ fault flag, TRUE when eErr is fault level
    bValid      : BOOL;  // 判定结果是否有效可用 ｜ check result valid flag
END_VAR
VAR
    bBad : BOOL; // 三输入非有限判定结果（NaN 或 ±Inf）｜ non-finite detection result of the three inputs
END_VAR

// 段 1｜返回值与输出预置 ｜ segment 1, preset return value and outputs
FC_DL_RangeCheckEx := FALSE; // 故障缺省判不在域内 ｜ fault default judges out-of-domain
bAboveUpper := FALSE;        // 预置未越上 ｜ preset not above upper
bBelowLower := FALSE;        // 预置未越下 ｜ preset not below lower
eErr        := 0;            // 预置无错误 ｜ preset no error
bError      := FALSE;        // 预置无故障 ｜ preset no fault
bValid      := FALSE;        // 预置无效，通过防御闸后置位 ｜ preset invalid, set TRUE after guard passes

// 段 2｜三输入非有限防御闸（早退） ｜ segment 2, non-finite guard of the three inputs (early return)
bBad := (fIn <> fIn) OR ((fIn - fIn) <> (fIn - fIn))
     OR (fLower <> fLower) OR ((fLower - fLower) <> (fLower - fLower))
     OR (fUpper <> fUpper) OR ((fUpper - fUpper) <> (fUpper - fUpper)); // 三输入非有限判定：NaN 自不等 + 差值自减判 ±Inf [无量纲] ｜ non-finite check: NaN by self-inequality, +/-Inf by self-subtraction
IF bBad THEN
    FC_DL_RangeCheckEx := FALSE; // 故障级判不在域内 ｜ fault level judges out-of-domain
    bAboveUpper := FALSE;        // 越上侧标志清零 ｜ clear the above-upper flag
    bBelowLower := FALSE;        // 越下侧标志清零 ｜ clear the below-lower flag
    eErr        := 16#0001_03CC; // 非有限输入故障码 ｜ non-finite input fault id
    bError      := TRUE;         // 置故障标志（R45 配对）｜ raise the fault flag (R45 pairing)
    bValid      := FALSE;        // 判定无效 ｜ check result invalid
    RETURN;                      // 早退 ｜ early return
END_IF

// 段 3｜双边界独立判定主体（末段） ｜ segment 3, independent per-boundary check body (final)
bAboveUpper := fIn > fUpper;  // 越上侧判定（与下限无关）｜ above-upper check (independent of the lower bound)
bBelowLower := fIn < fLower;  // 越下侧判定（与上限无关）｜ below-lower check (independent of the upper bound)
IF (NOT bAboveUpper) AND (NOT bBelowLower) THEN
    FC_DL_RangeCheckEx := TRUE;  // 双边界均未越，判在域内 ｜ neither boundary exceeded, judged in-domain
ELSE
    FC_DL_RangeCheckEx := FALSE; // 任一边界越出，判不在域内 ｜ either boundary exceeded, judged out-of-domain
END_IF
bError := FALSE; // 正常出口不置故障 ｜ normal exit raises no fault
bValid := TRUE;  // 判定输出有效可用 ｜ check output is valid
END_FUNCTION

(* ---- FC_DL_RatioToAmpDb.st ---- *)
(*
    FC_DL_RatioToAmpDb —— 线性幅值比到幅值型分贝换算
    ------------------------------------------------------------------
    分类      : DL_MathData / Log
    前缀      : FC_DL_
    版本      : 1.0.0
    溯源      : IEC 61131-3 标准语义的道莅防御性实现
                （接口语义由 IEC 61131-3 定义，内部委托平台内建 LOG，
                  外围统一错误码 / 钳位 / 双语文档；clean-room 重写，
                  未复制任何闭源厂商源码，参考实现仅限 MIT/Apache 许可）
    平台      : 纯 IEC 61131-3，CODESYS / TwinCAT / InoProShop 通用
    作者      : 道莅代码库 · PLC编程专家（R17）
    ------------------------------------------------------------------
    功能说明  : 线性幅值比转幅值型分贝值，按 dB = 20·log10(A) 实现，对数委托平台内建 LOG，
                20 为幅值型换算因子（与功率型 10 严格区分，禁混用），不重实现对数内核；
                非有限输入判为故障级 16#0001_02D3，返回 0.0 dB；
                定义域非法（比值 ≤ 0）判为故障级 16#0001_02D4，返回 0.0 dB；
                结果 |dB| 超 400.0 dB 时钳至 ±400.0 dB 并置信息级 16#0001_01EE
                （极小比值约 −760 dB，不钳会让下游 dB 域常量溢出）；
                钳位方向：结果双侧钳位至 ±400.0 dB。
    错误码    : 16#0001_01EE 结果超 ±400.0 dB，已钳至 dB 域硬限——信息级，正常防御
                16#0001_01EF 预留禁用（信息级，不得挪用）
                16#0001_02D3 非有限输入（NaN 或 ±INF）——故障级，返回 0.0
                16#0001_02D4 定义域非法（幅值比 ≤ 0）——故障级，返回 0.0
                16#0001_02D5 预留禁用（故障级，不得挪用）
    状态机    : R6 标注 N/A —— 本组件为纯函数无顺序状态机，无 CASE 可写，非法状态不可能出现，故以本节说明替代 ELSE 兜底
    修订记录  : 2026-11-16 v1.0.0 首次入库（R17）
*)
FUNCTION FC_DL_RatioToAmpDb : REAL
VAR_INPUT
    fRatio : REAL; // 线性幅值比（须 > 0，1.0 = 0 dB） [比] / linear amplitude ratio (must be > 0, 1.0 means 0 dB) [ratio]
END_VAR
VAR_OUTPUT
    eErr   : UDINT; // 错误码，0=正常 / error id, 0=ok
    bError : BOOL;  // 是否出错，eErr 非 0 时为 TRUE / error flag, TRUE when eErr is nonzero
    bValid : BOOL;  // 输出是否有效可用 / output valid flag
END_VAR
VAR CONSTANT
    DL_DB_FAULT_DEF   : REAL := 0.0;      // 故障缺省返回值（0 dB 中性值） [dB] / fault default return (0 dB neutral) [dB]
    DL_DB_AMP_FACTOR  : REAL := 20.0;     // 幅值型 dB 换算因子 20·log10 [dB] / amplitude dB factor 20*log10 [dB]
    DL_DB_LIMIT       : REAL := 400.0;    // dB 域双侧硬限 [dB] / two-sided dB hard limit [dB]
    DL_REAL_INF_GUARD : LREAL := 4.0E38;  // REAL 域 ±INF 判定阈值，高于 REAL 最大有限值 3.402823E38 [无量纲] / REAL +/-INF guard above max finite REAL
END_VAR
VAR
    fDb        : REAL; // dB 换算中间结果 [dB] / intermediate dB result [dB]
    bNonFinite : BOOL; // 非有限（NaN 或 ±INF）判定结果 / non-finite (NaN or +/-INF) detection result
END_VAR

// 段 1｜返回值与错误状态预置 / segment 1, preset return value and error status
FC_DL_RatioToAmpDb := DL_DB_FAULT_DEF; // 故障缺省返回 0 dB 中性值 [dB] / fault default 0 dB neutral value [dB]
eErr   := 0;     // 预置无错误 / preset no error
bError := FALSE; // 预置无故障 / preset no fault
bValid := FALSE; // 预置输出无效，通过全部域门后置位 / preset invalid, set TRUE after all domain gates

// 段 2｜非有限防御闸 / segment 2, non-finite guard
bNonFinite := (fRatio <> fRatio) OR (fRatio > DL_REAL_INF_GUARD) OR (fRatio < -DL_REAL_INF_GUARD); // 非有限判定（NaN 自不等 + 安全幅值判 ±INF） [比] / non-finite check (NaN by self-inequality, +/-INF by safe magnitude) [ratio]
IF bNonFinite THEN
    eErr := 16#0001_02D3; // 非有限输入故障码 / non-finite input fault id
    bError := TRUE;       // 置故障标志 / raise error flag
    bValid := FALSE;      // 输出不可用 / output not usable
    RETURN;               // 故障级提前返回，保持缺省 0 dB / early return on fault, keep default 0 dB
END_IF

// 段 3｜定义域（域门）判定 / segment 3, domain gate
IF fRatio <= 0.0 THEN
    eErr := 16#0001_02D4; // 定义域非法故障码（比值 ≤ 0，零点与负数无对数） [比] / domain fault id, ratio <= 0 has no logarithm [ratio]
    bError := TRUE;       // 置故障标志 / raise error flag
    bValid := FALSE;      // 输出不可用 / output not usable
    RETURN;               // 故障级提前返回，保持缺省 0 dB / early return on fault, keep default 0 dB
END_IF

// 段 4｜主体对数换算与结果钳位（末段） / segment 4, main logarithm conversion and result clamp (final)
fDb := LOG(fRatio) * DL_DB_AMP_FACTOR; // 委托内建 LOG 后乘幅值型因子 20 [dB] / delegate to built-in LOG then multiply amplitude factor 20 [dB]
IF fDb > DL_DB_LIMIT THEN
    fDb := DL_DB_LIMIT;   // 上侧钳至 +400.0 dB [dB] / clamp upward to +400.0 dB [dB]
    eErr := 16#0001_01EE; // 信息级：结果超硬限已钳位，正常防御 / info level: result exceeded the hard limit and was clamped
ELSIF fDb < -DL_DB_LIMIT THEN
    fDb := -DL_DB_LIMIT;  // 下侧钳至 −400.0 dB（极小比值不钳会使下游常量溢出） [dB] / clamp downward to -400.0 dB, tiny ratios would overflow downstream constants [dB]
    eErr := 16#0001_01EE; // 同一业务语义复用同一信息码 / same business semantics reuses the same info id
ELSE
    eErr := 0;            // 域内无错误 / in-domain, no error
END_IF
FC_DL_RatioToAmpDb := fDb; // 输出钳位后的 dB 结果 [dB] / output the clamped dB result [dB]
bError := FALSE;           // 信息级不置故障 / info level never raises fault
bValid := TRUE;            // 域内或钳位后输出均有效可用 / in-domain or clamped output is valid
END_FUNCTION

(* ---- FC_DL_RatioToPwrDb.st ---- *)
(*
    FC_DL_RatioToPwrDb —— 功率比值到 dB（10 因子）
    ------------------------------------------------------------------
    分类      : DL_MathData / Convert
    前缀      : FC_DL_
    版本      : 1.0.0
    溯源      : dB 为公开工程约定（功率型 10·log10，幅值型 20·log10）；本件为
                R17 件 FC_DL_PwrDbToRatio 的严格逆运算，补齐「功率型反向」缺位；
                定义域闸、零功率下限替代、饱和限与错误分级 100% 自有；
                对数一律委托平台内建 LN 换底，禁多项式重实现（T0 判据 2）；
                clean-room 重写，未复制任何闭源厂商源码，参考实现仅限 MIT/Apache 许可
    平台      : 纯 IEC 61131-3，CODESYS V3.5+ / TwinCAT 3 / InoProShop 通用
    作者      : 道莅代码库 · PLC编程专家（R19）
    ------------------------------------------------------------------
    功能说明  : 把功率比值报成 dB，用于射频电源、加热功率、光伏组串失配损耗的查表回算。
                核心防御：① fP2 ≤ 0 或 fP1 < 0 是定义域闸（负功率表示方向而非幅值，
                   比值语义失效），故障级 0324 早退；
                ② fP1 = 0 时按数学真值应为 -∞，本件在取对数之前就走定义域闸，
                   直接输出 fDbFloor（工程替代值）+ 信息 0404，绝不让 -∞ 出现；
                ③ 结果超 ±fDbSpan 双侧钳位，禁 NaN / ±INF 穿透；
                ④ 饱和硬限 380 dB 的可表性反算：380 dB → 10^38 < LREAL 上限，可表；
                   400 dB → 10^40 在 REAL 域不可表，故上限取 380 dB（R63 口径）。
                职责边界：本件只做比值→dB，正向换算归 FC_DL_PwrDbToRatio；参数超域按
                VAR CONSTANT 域钳位，钳位本身不置码（0405 只表结果超 span）。
    错误码    : 16#0001_0404 fP1 = 0，已按 fDbFloor 输出（真 -∞ 的工程替代）——信息级，正常防御
                16#0001_0405 结果超 ±fDbSpan 已钳位（bSaturated = TRUE）——信息级，正常防御
                16#0001_0324 功率非法（fP2 ≤ 0 或 fP1 < 0）——故障级，返回 0.0 且 bValid = FALSE
                16#0001_0325 输入或中间结果非有限（NaN / ±INF）——故障级，返回 0.0
                16#0001_0326 预留禁用（故障级，不得挪用）
    码位总账  : 16#0001_0404 用 / 16#0001_0405 用 ｜ 16#0001_0324 用 / 16#0001_0325 用 / 16#0001_0326 预留
    状态机    : R6 标注 N/A —— 本组件为纯函数无顺序状态机，无 CASE 可写，非法状态不可能出现
    采样约定  : 本件无定时器、无沿检测、无状态；单拍纯计算，结论与任务周期无关。
    修订记录  : 2026-11-16 v1.0.0 首次入库（R19）
*)
FUNCTION FC_DL_RatioToPwrDb : LREAL
VAR_INPUT
    fP1             : LREAL := 1.0;           // 分子功率 [W]，域 0.0~1.0E30，0 合法 / numerator power [W], range 0.0~1.0E30, zero allowed
    fP2             : LREAL := 1.0;           // 分母功率（参考功率）[W]，必须 > 0 / denominator reference power [W], must be > 0
    fDbSpan         : LREAL := 380.0;         // dB 绝对值上限 [dB]，域 1.0~1000.0 / absolute dB span [dB], range 1.0~1000.0
    fDbFloor        : LREAL := -380.0;        // fP1 = 0 时的下限替代值 [dB]，域 -1000.0~0.0 / floor substitute when fP1 = 0 [dB], range -1000.0~0.0
END_VAR
VAR_OUTPUT
    eErr            : UDINT;                  // 错误码，0=正常 / error id, 0=ok
    bError          : BOOL;                   // 故障标志，eErr 为故障级时 TRUE / error flag, TRUE on fault-level eErr
    bValid          : BOOL;                   // 返回值是否可用 / return value valid flag
    bSaturated      : BOOL;                   // 结果被钳位 / result clamped
    bZeroPower      : BOOL;                   // fP1 = 0，真 -∞ 已按下限替代 / fP1 = 0, true minus infinity replaced by the floor
END_VAR
VAR CONSTANT
    DL_DB_PWR_FACTOR : LREAL := 10.0;         // 功率型 dB 因子 [无量纲] / power dB factor [dimensionless]
    DL_LOG_BASE10    : LREAL := 10.0;         // 换底用对数的底 [无量纲] / logarithm base for the base change [dimensionless]
    DL_FLOAT_EPS     : REAL := 1.0E-6;        // 浮点判等容差 [无量纲] / float equality tolerance [dimensionless]
    DL_DB_SPAN_MIN   : LREAL := 1.0;          // dB 上限最小值 [dB] / minimum dB span [dB]
    DL_DB_SPAN_MAX   : LREAL := 1000.0;       // dB 上限最大值 [dB] / maximum dB span [dB]
    DL_DB_FLOOR_MIN  : LREAL := -1000.0;      // 下限替代值最小值 [dB] / minimum floor substitute [dB]
    DL_DB_FLOOR_MAX  : LREAL := 0.0;          // 下限替代值最大值 [dB] / maximum floor substitute [dB]
    DL_DB_INF_GUARD  : LREAL := 1.0E300;      // 非有限幅值判定阈值 [无量纲] / non-finite magnitude guard [dimensionless]
    DL_DB_ZERO       : LREAL := 0.0;          // 零值常量，避免裸字面量 [dB] / zero constant, avoids a bare literal [dB]
END_VAR
VAR
    fRatio          : LREAL;                  // 功率比值 fP1/fP2 [无量纲] / power ratio fP1/fP2 [dimensionless]
    fDb             : LREAL;                  // 计算中的 dB 中间量 [dB] / dB intermediate value [dB]
    fSpanEff        : LREAL;                  // 生效 dB 上限，域钳位后使用 [dB] / effective dB span after clamping [dB]
    fFloorEff       : LREAL;                  // 生效下限替代值，域钳位后使用 [dB] / effective floor substitute after clamping [dB]
    bNonFin         : BOOL;                   // 输入非有限判定标志 / non-finite input flag
END_VAR

// 段 1｜返回值与错误状态预置 / segment 1, preset return value and error status
FC_DL_RatioToPwrDb := DL_DB_ZERO;             // 故障缺省返回 0 dB / fault default returns zero dB
eErr := 0;                                    // 预置无错误 / preset no error
bError := FALSE;                              // 预置无故障 / preset no fault
bValid := FALSE;                              // 预置不可用，通过闸门后置位 / preset invalid, set TRUE after the gates
bSaturated := FALSE;                          // 预置未饱和 / preset not saturated
bZeroPower := FALSE;                          // 预置非零功率 / preset non-zero power

// 段 2｜非有限输入闸（NaN 穿透拦截，先于任何比较与对数）/ segment 2, non-finite input gate
bNonFin := (fP1 <> fP1) OR (fP1 > DL_DB_INF_GUARD) OR (fP1 < -DL_DB_INF_GUARD)
        OR (fP2 <> fP2) OR (fP2 > DL_DB_INF_GUARD) OR (fP2 < -DL_DB_INF_GUARD)
        OR (fDbSpan <> fDbSpan) OR (fDbFloor <> fDbFloor);  // 非有限判定 / non-finite detection
IF bNonFin THEN
    eErr := 16#0001_0325;                     // 输入非有限故障码 / non-finite input fault id
    bError := TRUE;                           // 置故障标志 / raise the error flag
    RETURN;                                   // 故障级提前返回 / early return on fault
END_IF

// 段 3｜定义域闸：分母非正、分子为负均为非法功率语义 / segment 3, domain gate on the powers
IF (fP2 <= DL_DB_ZERO) OR (fP1 < DL_DB_ZERO) THEN
    eErr := 16#0001_0324;                     // 功率非法故障码 / illegal power fault id
    bError := TRUE;                           // 置故障标志 / raise the error flag
    RETURN;                                   // 故障级提前返回，绝不进入对数 / early return, the logarithm is never executed
END_IF

// 段 4｜参数域钳位（上限、下限替代值各自双侧收敛，钳位本身不置码）/ segment 4, parameter domain clamp
fSpanEff := MIN(MAX(fDbSpan, DL_DB_SPAN_MIN), DL_DB_SPAN_MAX);     // 上限收敛到 1.0~1000.0 dB / converge the span into 1.0~1000.0 dB
fFloorEff := MIN(MAX(fDbFloor, DL_DB_FLOOR_MIN), DL_DB_FLOOR_MAX); // 下限替代收敛到 -1000.0~0.0 dB / converge the floor into -1000.0~0.0 dB

// 段 5｜零功率闸：定义域闸优于事后判 -∞，直接给工程替代值 / segment 5, zero power gate
IF ABS(fP1) <= DL_FLOAT_EPS THEN
    bZeroPower := TRUE;                       // 标记零功率 / flag the zero power
    bValid := TRUE;                           // 替代值可用 / the substitute is usable
    eErr := 16#0001_0404;                     // 信息级：真 -∞ 的工程替代 / info level, engineering substitute for minus infinity
    IF fFloorEff > -fSpanEff THEN
        FC_DL_RatioToPwrDb := fFloorEff;      // 下限未越 span 时按入参输出 / publish the floor when it stays inside the span
    ELSE
        FC_DL_RatioToPwrDb := -fSpanEff;      // 下限越 span 时钳到 -span，保持双侧一致 / clamp to minus span to keep both sides consistent
        bSaturated := TRUE;                   // 标记饱和 / flag the saturation
    END_IF
    RETURN;                                   // 零功率分支出口，不取对数 / exit without taking any logarithm
END_IF

// 段 6｜委托内建 LN 换底（禁多项式重实现）/ segment 6, delegate to the built-in LN with a base change
fRatio := fP1 / fP2;                          // 分母已由段 3 保证 > 0，除法安全 / the denominator is positive by segment 3, the division is safe
fDb := DL_DB_PWR_FACTOR * (LN(fRatio) / LN(DL_LOG_BASE10)); // 10·log10(P1/P2) / 10 log10 of the power ratio

// 段 7｜结果非有限复检 / segment 7, non-finite recheck
IF (fDb <> fDb) OR (fDb > DL_DB_INF_GUARD) OR (fDb < -DL_DB_INF_GUARD) THEN
    eErr := 16#0001_0325;                     // 中间结果非有限故障码 / non-finite intermediate fault id
    bError := TRUE;                           // 置故障标志 / raise the error flag
    FC_DL_RatioToPwrDb := DL_DB_ZERO;         // 明确返回 0 dB / return zero dB explicitly
    RETURN;                                   // 故障级提前返回 / early return on fault
END_IF

// 段 8｜双侧饱和钳位 / segment 8, two-sided saturation clamp
IF fDb > fSpanEff THEN
    fDb := fSpanEff;                          // 正向超限钳位 / clamp the positive overrun
    bSaturated := TRUE;                       // 标记饱和 / flag the saturation
    eErr := 16#0001_0405;                     // 信息级：超 span 已钳位 / info level, clamped to the span
ELSIF fDb < -fSpanEff THEN
    fDb := -fSpanEff;                         // 负向超限钳位 / clamp the negative overrun
    bSaturated := TRUE;                       // 标记饱和 / flag the saturation
    eErr := 16#0001_0405;                     // 同一业务语义复用同一信息码 / the same semantics reuses the same info id
END_IF

// 段 9｜发布结果 / segment 9, publish the result
FC_DL_RatioToPwrDb := fDb;                    // 输出 dB 值 [dB] / publish the dB value [dB]
bValid := TRUE;                               // 通过全部闸门，结果可用 / all gates passed, the result is usable
bError := FALSE;                              // 信息级不置故障 / info level never raises a fault
END_FUNCTION

(* ---- FC_DL_RealEqTolEx.st ---- *)
(*
    FC_DL_RealEqTolEx —— 浮点容差判等原子（LREAL 域）
    ------------------------------------------------------------------
    分类      : DL_MathData / Compare
    前缀      : FC_DL_
    版本      : 1.0.0
    溯源      : IEC 61131-3 标准语义的道莅防御性实现
                （内部委托 ABS 标准运算与比较语义，外围统一错误码/钳位/双语文档；
                  未复制任何闭源厂商源码，参考实现仅限 MIT/Apache 许可）
    平台      : 纯 IEC 61131-3，CODESYS / TwinCAT / InoProShop 通用
    作者      : 道莅代码库 · PLC编程专家（R40）
    ------------------------------------------------------------------
    功能说明  : 浮点容差判等原子：当 ABS(fA − fB) ≤ fTol 时判为相等（含边界，
                「差值不超过容差」即视为相等，全库口径统一按本件为准）；
                本件为红线 5「浮点判等禁用 = / <>」的库级原子化出口，
                全库判等口径以引用本件为准（语义引用，不强制实例化调用）；
                任一输入非有限（NaN 或 ±Inf）判为故障级 16#0001_03CB，
                返回 FALSE 且 bValid=FALSE（NaN 与任何值比较均无意义，一律拦截）；
                非有限判定口径（R15）：NaN 用自不等 f <> f，±Inf 用 (f − f) <> (f − f)；
                容差下限防死判：fTol 有限但小于容差下限 1.0E-9（含负值与 0）时
                钳至下限并置信息级 16#0001_0492——容差为 0 或近 0 会使判等恒 FALSE
                （浮点差值几乎不可能精确为 0，形成「死判」），下限钳位保证判等可用。
    错误码    : 16#0001_03CB 任一输入非有限（NaN 或 ±Inf）——故障级，返回 FALSE
                16#0001_0492 容差小于下限 1.0E-9（含负值与 0），已钳至下限——信息级，正常防御
                （R90 反证句：容差被钳这一事实无法由返回值观测——返回 TRUE 与 FALSE
                  均可能在钳位前后同时出现，现有输出组合无法还原「容差已被钳」场景，故占信息码）
    状态机    : R6 标注 N/A —— 本组件为纯函数无顺序状态机，无 CASE 可写，
                非法状态不可能出现，故以本节说明替代 ELSE 兜底
    修订记录  : 2026-11-19 v1.0.0 首次入库（R40 · 批 1 · T0 快车道）
*)
FUNCTION FC_DL_RealEqTolEx : BOOL
VAR_INPUT
    fA   : LREAL; // 比较左值 [无量纲] ｜ left comparand
    fB   : LREAL; // 比较右值 [无量纲] ｜ right comparand
    fTol : LREAL; // 容差 [无量纲]，小于下限或非正时钳至下限 ｜ tolerance, clamped to the floor when below it or non-positive
END_VAR
VAR_OUTPUT
    eErr   : UDINT; // 错误码，0=正常，16#0001_04XX=信息级，16#0001_03XX=故障级 ｜ error id, 0=ok, 16#0001_04XX=info, 16#0001_03XX=fault
    bError : BOOL;  // 是否出错，eErr 落故障级时为 TRUE ｜ fault flag, TRUE when eErr is fault level
    bValid : BOOL;  // 输出是否有效可用 ｜ output valid flag
END_VAR
VAR CONSTANT
    DL_TOL_FLOOR : LREAL := 1.0E-9; // 容差下限，防止零容差死判 [无量纲] ｜ tolerance floor, prevents the zero-tolerance dead comparison
END_VAR
VAR
    bBad    : BOOL;  // 三输入非有限判定结果（NaN 或 ±Inf）｜ non-finite detection result of the three inputs
    fTolEff : LREAL; // 整备后的有效容差 [无量纲] ｜ effective tolerance after preparation
    fDiff   : LREAL; // 两值差值绝对值 [无量纲] ｜ absolute difference of the two values
END_VAR

// 段 1｜返回值与错误状态预置 ｜ segment 1, preset return value and error status
FC_DL_RealEqTolEx := FALSE; // 故障缺省返回不相等 ｜ fault default returns not-equal
eErr   := 0;     // 预置无错误 ｜ preset no error
bError := FALSE; // 预置无故障 ｜ preset no fault
bValid := FALSE; // 预置无效，通过防御闸后置位 ｜ preset invalid, set TRUE after guard passes

// 段 2｜三输入非有限防御闸（早退） ｜ segment 2, non-finite guard of the three inputs (early return)
bBad := (fA <> fA) OR ((fA - fA) <> (fA - fA))
     OR (fB <> fB) OR ((fB - fB) <> (fB - fB))
     OR (fTol <> fTol) OR ((fTol - fTol) <> (fTol - fTol)); // 三输入非有限判定：NaN 自不等 + 差值自减判 ±Inf [无量纲] ｜ non-finite check: NaN by self-inequality, +/-Inf by self-subtraction
IF bBad THEN
    FC_DL_RealEqTolEx := FALSE; // 故障级返回不相等 ｜ fault level returns not-equal
    eErr   := 16#0001_03CB;     // 非有限输入故障码 ｜ non-finite input fault id
    bError := TRUE;             // 置故障标志（R45 配对）｜ raise the fault flag (R45 pairing)
    bValid := FALSE;            // 输出无效 ｜ output invalid
    RETURN;                     // 早退 ｜ early return
END_IF

// 段 3｜容差下限钳位（防死判） ｜ segment 3, tolerance floor clamp (prevents the dead comparison)
IF fTol < DL_TOL_FLOOR THEN
    fTolEff := DL_TOL_FLOOR; // 容差钳至下限 [无量纲] ｜ tolerance clamped to the floor
    eErr    := 16#0001_0492; // 信息级：容差已钳下限 ｜ info level: tolerance clamped to the floor
ELSE
    fTolEff := fTol;         // 域内容差直通 [无量纲] ｜ in-domain tolerance pass-through
END_IF

// 段 4｜容差判等主体（末段） ｜ segment 4, tolerance equality body (final)
fDiff := ABS(fA - fB);       // 差值绝对值 [无量纲] ｜ absolute difference
IF fDiff <= fTolEff THEN
    FC_DL_RealEqTolEx := TRUE;  // 差值不超过有效容差，判相等（含边界）｜ difference within the effective tolerance, judged equal (boundary inclusive)
ELSE
    FC_DL_RealEqTolEx := FALSE; // 差值超容差，判不等 ｜ difference beyond the tolerance, judged not-equal
END_IF
bError := FALSE; // 信息级钳位不置故障，故障分支已提前返回 ｜ info-level clamp never raises fault, fault branch has returned
bValid := TRUE;  // 判等输出有效可用 ｜ comparison output is valid
END_FUNCTION

(* ---- FC_DL_RealToByteSat.st ---- *)
(*
    FC_DL_RealToByteSat —— REAL 到 BYTE 饱和防御转换
    ------------------------------------------------------------------
    分类      : DL_MathData / Convert
    前缀      : FC_DL_
    版本      : 1.0.0
    溯源      : IEC 61131-3 标准语义的道莅防御性实现
                （内部委托平台内建函数，外围统一错误码/钳位/双语文档；
                  未复制任何闭源厂商源码，参考实现仅限 MIT/Apache 许可）
    平台      : 纯 IEC 61131-3，CODESYS / TwinCAT / InoProShop 通用
    作者      : 道莅代码库 · PLC编程专家（R16）
    ------------------------------------------------------------------
    功能说明  : 将 REAL 输入防御性转换为 BYTE 并作为返回值输出，面向串口报文字节域
                与 PWM 占空比字节域（0~255）等单字节输出场景；
                非有限输入（NaN 或 ±INF）判为故障级 16#0001_029A，返回 0 且 bValid=FALSE；
                fIn < 0 时钳位至 0，置信息级 16#0001_01C8（BYTE 无符号，负值不可表）；
                fIn 超出 BYTE 上界 255 时钳位至上界，置信息级 16#0001_01C9（串口/PWM 占空比字节域用途）；
                钳位方向：下界 0 / 上界 255（双侧饱和）；
                ±INF 采用平台安全幅值比较判定（阈值高于 REAL 最大有限值 3.402823E38），NaN 用 fIn <> fIn 自不等判定；
                域内转换委托平台内建 REAL_TO_BYTE 语义，不重实现数学内核；
                信息级码属正常防御：bError=FALSE、bValid=TRUE，输出钳位后防御值。
    错误码    : 16#0001_029A 非有限输入（NaN 或 ±INF）——故障级，返回 0
                16#0001_01C8 负值输入，已钳位至 0——信息级，正常防御
                16#0001_01C9 输入超 BYTE 上界，已钳位至 255——信息级，正常防御
                16#0001_029B 预留禁用（故障级，不得挪用）
                16#0001_029C 预留禁用（故障级，不得挪用）
    状态机    : R6 标注 N/A —— 本组件为纯函数无顺序状态机，无 CASE 可写，非法状态不可能出现，故以本节说明替代 ELSE 兜底
    修订记录  : 2026-11-16 v1.0.0 首次入库（R16）
*)
FUNCTION FC_DL_RealToByteSat : BYTE
VAR_INPUT
    fIn : REAL; // 待转换输入 [无量纲] / input value to convert
END_VAR
VAR_OUTPUT
    eErr   : UDINT; // 错误码，0=正常 / error id, 0=ok
    bError : BOOL;  // 是否出错，eErr 非 0 时为 TRUE / error flag, TRUE when eErr is nonzero
    bValid : BOOL;  // 输出是否有效可用 / output valid flag
END_VAR
VAR CONSTANT
    DL_BYTE_MAX       : LREAL := 255.0; // BYTE 域上界 255，LREAL 承载 [无量纲] / BYTE upper bound 255 carried in LREAL
    DL_REAL_INF_GUARD : LREAL := 4.0E38; // REAL 域 ±INF 判定阈值，高于 REAL 最大有限值 3.402823E38 [无量纲] / REAL +/-INF guard above max finite REAL 3.402823E38
END_VAR
VAR
    bNonFinite : BOOL; // 非有限（NaN 或 ±INF）判定结果 / non-finite (NaN or +/-INF) detection result
END_VAR

// 段 1｜返回值与错误状态预置 / segment 1, preset return value and error status
FC_DL_RealToByteSat := 16#00; // 故障缺省返回 0 [无量纲] / fault default returns 0
eErr   := 0;     // 预置无错误 / preset no error
bError := FALSE; // 预置无故障 / preset no fault
bValid := FALSE; // 预置无效，通过防御闸后置位 / preset invalid, set TRUE after guard passes

// 段 2｜非有限防御闸 / segment 2, non-finite guard
bNonFinite := (fIn <> fIn) OR (fIn > DL_REAL_INF_GUARD) OR (fIn < -DL_REAL_INF_GUARD); // NaN 自不等判定，±INF 用安全幅值比较 [无量纲] / NaN by self-inequality, +/-INF by safe magnitude compare
IF bNonFinite THEN
    FC_DL_RealToByteSat := 16#00; // 故障级返回 0 [无量纲] / fault level returns 0
    eErr   := 16#0001_029A;       // 非有限输入故障码 / non-finite input fault id
    bError := TRUE;               // 置故障标志 / set fault flag
    bValid := FALSE;              // 输出无效 / output invalid
    RETURN;                       // 立即返回 / immediate return
END_IF

// 段 3｜双侧饱和钳位与主体转换（末段） / segment 3, double-side saturating clamp and main conversion (final)
IF fIn < 0.0 THEN
    FC_DL_RealToByteSat := 16#00; // 负值钳位至 0（BYTE 无符号语义） / negative input clamped to 0 (BYTE is unsigned)
    eErr := 16#0001_01C8;         // 信息级：负值已钳零 / info level: negative input clamped to zero
ELSIF fIn > DL_BYTE_MAX THEN
    FC_DL_RealToByteSat := 16#FF; // 正向钳位至 BYTE 上界 255（串口/PWM 占空比字节域） / clamp to BYTE upper bound 255 (serial frame and PWM duty byte domain)
    eErr := 16#0001_01C9;         // 信息级：超上界已钳位 / info level: above upper bound, clamped
ELSE
    FC_DL_RealToByteSat := REAL_TO_BYTE(fIn); // 域内委托平台内建 _TO_ 转换语义 / in-domain delegate to built-in _TO_ conversion
    eErr := 0; // 域内无错误 / in-domain, no error
END_IF
bError := FALSE; // 信息级钳位不置故障，故障分支已提前返回 / info-level clamp never raises fault, fault branch has returned
bValid := TRUE;  // 域内或钳位输出均有效可用 / in-domain or clamped output is valid
END_FUNCTION

(* ---- FC_DL_RealToDintSat.st ---- *)
(*
    FC_DL_RealToDintSat —— LREAL/REAL 到 DINT 饱和防御降型
    ------------------------------------------------------------------
    分类      : DL_MathData / Convert
    前缀      : FC_DL_
    版本      : 1.0.0
    溯源      : IEC 61131-3 标准语义的道莅防御性实现
                （内部委托平台内建 LREAL_TO_DINT 转换语义，外围统一错误码/钳位/
                  双语文档；未复制任何闭源厂商源码，参考实现仅限 MIT/Apache 许可）
    平台      : 纯 IEC 61131-3，CODESYS / TwinCAT / InoProShop 通用
    作者      : 道莅代码库 · PLC编程专家（R40）
    ------------------------------------------------------------------
    功能说明  : 将 LREAL 输入（REAL 实参按标准隐式升位传入）防御性降型为 DINT
                并作为返回值输出，转换内核委托平台内建 LREAL_TO_DINT（向零截断），
                不重实现任何转换内核；
                非有限输入（NaN 或 ±Inf）判为故障级 16#0001_03CD，返回 0 且
                bValid=FALSE（非有限值参与降型在三平台行为不一致，一律拦截）；
                越界双侧显式钳位（R55/R241：跨类型降型禁靠隐式回绕兜底）：
                fIn > 2147483647.0 钳至 DINT 上界，置信息级 16#0001_0493；
                fIn < −2147483648.0 钳至 DINT 下界，置信息级 16#0001_0494；
                双侧直比判定，禁用 ABS 单侧判据（有符号最小值取 ABS 回绕会漏判）；
                转换前置域闸（先判域后转换）：域闸命中不调内建转换，
                保证 LREAL_TO_DINT 只接收域内可表值，杜绝降型溢出方向翻转；
                信息级码属正常防御：bError=FALSE、bValid=TRUE，输出钳位后防御值。
    错误码    : 16#0001_03CD 非有限输入（NaN 或 ±Inf）——故障级，返回 0
                16#0001_0493 输入超 DINT 上界 2147483647，已钳至上界——信息级，正常防御
                16#0001_0494 输入低于 DINT 下界 −2147483648，已钳至下界——信息级，正常防御
                （R90 反证句：越上界与越下界两场景均无法由返回值加 bValid 组合区分——
                  钳位后输出为合法边界值，bValid=TRUE 与域内转换相同，若共用一码则
                  现场无法还原越界方向，故两侧各占一码）
    非有限口径 : NaN 用自不等 f <> f，±Inf 用 (f − f) <> (f − f) 差值自减判定（R15）；
                LREAL 最大有限值之上无可表常量，禁用近似幅值阈值。
    状态机    : R6 标注 N/A —— 本组件为纯函数无顺序状态机，无 CASE 可写，
                非法状态不可能出现，故以本节说明替代 ELSE 兜底
    修订记录  : 2026-11-19 v1.0.0 首次入库（R40 · 批 2 · T0 快车道）
*)
FUNCTION FC_DL_RealToDintSat : DINT
VAR_INPUT
    fIn : LREAL; // 待降型输入 [无量纲]，REAL 实参按标准升位传入 ｜ input to down-convert, REAL arguments widen by standard rules
END_VAR
VAR_OUTPUT
    eErr   : UDINT; // 错误码，0=正常，16#0001_04XX=信息级，16#0001_03XX=故障级 ｜ error id, 0=ok, 16#0001_04XX=info, 16#0001_03XX=fault
    bError : BOOL;  // 是否出错，eErr 落故障级时为 TRUE ｜ fault flag, TRUE when eErr is fault level
    bValid : BOOL;  // 输出是否有效可用 ｜ output valid flag
END_VAR
VAR CONSTANT
    DL_DINT_MAX_R : LREAL := 2.147483647E9;  // DINT 上界 2147483647 的 LREAL 承载值 [无量纲] ｜ DINT upper bound 2147483647 carried in LREAL
    DL_DINT_MIN_R : LREAL := -2.147483648E9; // DINT 下界 −2147483648 的 LREAL 承载值 [无量纲] ｜ DINT lower bound −2147483648 carried in LREAL
END_VAR
VAR
    bNonFinite : BOOL; // 非有限（NaN 或 ±Inf）判定结果 ｜ non-finite (NaN or +/-Inf) detection result
END_VAR

// 段 1｜返回值与错误状态预置 ｜ segment 1, preset return value and error status
FC_DL_RealToDintSat := 0; // 故障缺省返回 0 [无量纲] ｜ fault default returns 0
eErr   := 0;     // 预置无错误 ｜ preset no error
bError := FALSE; // 预置无故障 ｜ preset no fault
bValid := FALSE; // 预置无效，通过防御闸后置位 ｜ preset invalid, set TRUE after guard passes

// 段 2｜非有限防御闸（命中不调内建转换，早退） ｜ segment 2, non-finite guard (early return, no built-in conversion)
bNonFinite := (fIn <> fIn) OR ((fIn - fIn) <> (fIn - fIn)); // NaN 自不等 + 差值自减判 ±Inf [无量纲] ｜ NaN by self-inequality, +/-Inf by self-subtraction
IF bNonFinite THEN
    FC_DL_RealToDintSat := 0; // 故障级返回 0 [无量纲] ｜ fault level returns 0
    eErr   := 16#0001_03CD;   // 非有限输入故障码 ｜ non-finite input fault id
    bError := TRUE;           // 置故障标志（R45 配对）｜ raise the fault flag (R45 pairing)
    bValid := FALSE;          // 输出无效 ｜ output invalid
    RETURN;                   // 早退，不调内建转换 ｜ early return, no built-in conversion
END_IF

// 段 3｜越界双侧显式钳位与域内转换（末段，先判域后转换） ｜ segment 3, double-side explicit clamp and in-domain conversion (final, domain check before conversion)
IF fIn > DL_DINT_MAX_R THEN
    FC_DL_RealToDintSat := 2147483647;  // 越上界钳至 DINT 上界 [无量纲] ｜ above upper bound, clamp to the DINT upper bound
    eErr := 16#0001_0493;               // 信息级：越上界已钳位 ｜ info level: above upper bound, clamped
ELSIF fIn < DL_DINT_MIN_R THEN
    FC_DL_RealToDintSat := -2147483648; // 越下界钳至 DINT 下界 [无量纲] ｜ under lower bound, clamp to the DINT lower bound
    eErr := 16#0001_0494;               // 信息级：越下界已钳位 ｜ info level: under lower bound, clamped
ELSE
    FC_DL_RealToDintSat := LREAL_TO_DINT(fIn); // 域内委托平台内建降型转换（向零截断）｜ in-domain delegate to the built-in down-conversion (truncate toward zero)
    eErr := 0;                                 // 域内无错误 ｜ in-domain, no error
END_IF
bError := FALSE; // 信息级钳位不置故障，故障分支已提前返回 ｜ info-level clamp never raises fault, fault branch has returned
bValid := TRUE;  // 域内或钳位输出均有效可用 ｜ in-domain or clamped output is valid
END_FUNCTION

(* ---- FC_DL_RealToIntSat.st ---- *)
(*
  ==================================================================
  组件名 Component  : FC_DL_RealToIntSat
  分类   Category   : DL_MathData
  前缀   Naming     : FC_DL_ ｜ b/n/u/f/t/e/st 类型前缀制（R265）
  码位   Code ID    : 16#0001_064E（信息级）｜ 16#0001_064F / 0650（故障级）
  版本   Version    : 1.0.0
  复杂度 Complexity  : 中
  功能   Purpose    : LREAL → INT（16 位）饱和转换，统一三平台「部分平台饱和、部分平台
                      回绕」的差异；NaN / ±Inf / 越界全部确定性处置。
  开源溯源 Origin    : IEC 61131-3 标准语义的道莅防御性实现（clean-room，无第三方代码行）
  许可证 License    : MIT
  参考   Reference  : IEC 61131-3:2013 §6.6.5 类型转换函数（REAL 到整型的截断语义）
  平台   Platform   : 纯 IEC 61131-3（LREAL_TO_INT / 比较），三平台通用
  依赖   Depends    : 仅 Standard.library（LREAL_TO_INT 属标准转换函数）
  分工声明 Split     : FC_DL_RealToDintSat（32 位）与 FC_DL_RealToByteSat（8 位）为同位宽
                      兄弟件，本件补 INT（16 位），三件构成位宽三分（R216 双向互引）；
                      工程舍入（四舍五入）归 FC_DL_RoundSat，有效位舍入归 FC_DL_RoundSigFigs，
                      本件只做向零截断。
  归属 Ownership     : 本件无 TYPE 声明，全部引脚为 IEC 标准原生类型。
  编译门槛 Gate      : 交付门槛：主路径委托平台内建 LREAL_TO_INT，其截断（向零）语义须在
                      CODESYS / TwinCAT 3 / InoProShop 三平台各编译并跑一次本文件 V2 向量
                      （R64 内建转换链交付门槛）。
  ------------------------------------------------------------------
  边界 Boundary     :
                      一 判据严格有序：① NaN → 0 + 故障码 + bValid FALSE + 早退；
                         ② 组态 nLo > nHi → 故障码 + 早退；③ ±Inf → 对应边界；
                         ④ 越界 → 钳边界 + bClamped；⑤ 域内 → 向零截断；
                      二 一律在转换之前做域钳（R151：实数转整数前先钳，防溢出使方向翻转）；
                      三 非有限判据用自反与差值自减，禁用近似阈值（R79）：
                         NaN 用 fIn <> fIn，Inf 用 (fIn − fIn) <> (fIn − fIn)；
                      四 bClamped 与 bNonFinite 语义可分：域钳只置前者，非有限两者都置；
                      五 nLo > nHi 判组态故障返回 FALSE（与 FC_DL_SaturateMul / Div 同口径）；
                      六 纯函数：无记忆量、无定时器、无边沿实例，每调用重算。
  错误码 Codes      :
    16#0001_064E【信息级】输入越 [nLo, nHi] 已钳边界（bClamped = TRUE，bValid = TRUE）
    16#0001_064F【故障级】输入非有限（NaN 返 0；±Inf 钳对应边界；bValid = FALSE）
    16#0001_0650【故障级】组态非法 nLo > nHi（判故障返回 FALSE，nOut = 0）
  码位反证 Note     :
    064E 不可并入 064F：域钳结果可用（bValid = TRUE、无 bError），非有限结果不可用，
    上游 HMI 按 bValid 过滤时两者必须分开，合并会让「钳位可用」被当成「测点坏」停机（R90）。
  验收 Acceptance   :
    算法已证（脚本）：未跑 ｜ 编译器已证（三平台）：未跑
    V1 0.0 → 0、bClamped = FALSE、无码
    V2 -0.5 → 0（向零截断）、bClamped = FALSE（域内，仅截断）
    V3 32767.9 → 32767（越上界半个 LSB，钳上界）
    V4 32768.0 → 32767 + bClamped + 码 064E
    V5 -32768.1 → -32768 + bClamped + 码 064E
    V6 NaN → 0 + bNonFinite = TRUE + bValid = FALSE + 码 064F
    V7 1.0E9 → 32767 + bClamped + 码 064E
    V8 nLo > nHi → 码 0650 + 返回 FALSE
    V9 nLo = nHi = 100 → 恒定输出 100 + bClamped（域退化）
  修订记录 Revision  :
    2026-11-21  v1.0.0  R62 首版（批 2 · 序号 5）
  ==================================================================
*)
FUNCTION FC_DL_RealToIntSat : BOOL
VAR_INPUT
    fIn : LREAL;          // 输入量 [工程单位]，必须有限 / the input value, must be finite
    nLo : INT := -32768;  // 目标钳位域下界 [−]，默认 INT 全域下界 / the clamp floor, the INT domain floor by default
    nHi : INT := 32767;   // 目标钳位域上界 [−]，默认 INT 全域上界 / the clamp ceiling, the INT domain ceiling by default
END_VAR
VAR_OUTPUT
    nOut      : INT;   // 饱和转换结果 [−] / the saturated integer result
    bClamped  : BOOL;  // 域钳位发生（含 ±Inf 钳边界）[-] / a domain clamp happened, the infinite boundary clamp included
    bNonFinite: BOOL;  // 输入非有限（NaN 或 ±Inf）[-] / the input was not finite
    bValid    : BOOL;  // 输出可用（非有限与组态故障为 FALSE）[-] / the output is usable
    eErr      : UDINT; // 错误码，0 = 正常 / the error code, zero is ok
    bError    : BOOL;  // 故障标志，故障级码同拍置位（R45 配对）/ the fault flag, raised with a fault level code
END_VAR
VAR
    fLo : LREAL := 0.0; // 下界的实数形式 [−] / the floor in real form
    fHi : LREAL := 0.0; // 上界的实数形式 [−] / the ceiling in real form
END_VAR  // R64 结构补齐：VAR 段缺失的 END_VAR（门禁机械修复）
VAR CONSTANT
    DL_R2I_ZERO : LREAL := 0.0;   // 实数零常量 [−] / the real zero constant
    DL_R2I_NONE : INT := 0;       // 整型零常量 [−] / the integer zero constant
END_VAR

// 段 1｜返回值与全部出口预置安全值（R45 四段式第一段）/ segment 1, preset every outlet to its safe value
FC_DL_RealToIntSat := FALSE; // 返回值预置假 / preset the return false
nOut := DL_R2I_NONE; // 结果预置零 [−] / preset the result zero
bClamped := FALSE; // 钳位标志预置假 / preset the clamp flag false
bNonFinite := FALSE; // 非有限标志预置假 / preset the non finite flag false
bValid := FALSE; // 可用标志预置假，过闸后置位 / preset the validity false, raised after the gates
eErr := 16#0000_0000; // 错误码预置正常 / preset the code to ok
bError := FALSE; // 故障标志预置假 / preset the fault flag false
fLo := DL_R2I_ZERO; // 下界实数形式清零 / clear the floor in real form
fHi := DL_R2I_ZERO; // 上界实数形式清零 / clear the ceiling in real form

// 段 2｜判据①NaN：自反性判定，禁近似阈值（边界三，R79）/ segment 2, the NaN gate by reflexivity
IF fIn <> fIn THEN // NaN：一切比较均为假，只能用自反性 / NaN leaves every comparison false, reflexivity is the only test
    bNonFinite := TRUE; // 置非有限标志 / raise the non finite flag
    bValid := FALSE; // 结果不可用（三件套之一，R258）/ the result is not usable
    nOut := DL_R2I_NONE; // 确定缺省值零 [−] / the deterministic default of zero
    eErr := 16#0001_064F; // 故障级：输入非有限 / fault grade, the input is not finite
    bError := TRUE; // 同拍置故障标志（R45 配对）/ raise the fault flag on the same scan
    RETURN; // 早退 / early return
END_IF

// 段 3｜判据②组态域闸：nLo > nHi 判故障早退（边界五）/ segment 3, the configuration gate, a reversed domain is a fault
IF nLo > nHi THEN // 钳位域反序 / the clamp domain is reversed
    eErr := 16#0001_0650; // 故障级：组态非法 nLo > nHi / fault grade, the reversed clamp domain
    bError := TRUE; // 同拍置故障标志（R45 配对）/ raise the fault flag on the same scan
    bValid := FALSE; // 输出不可用 / the output is not usable
    nOut := DL_R2I_NONE; // 确定缺省值零 [−] / the deterministic default of zero
    RETURN; // 早退 / early return
END_IF

// 段 4｜判据③±Inf：差值自减判无穷（边界三），钳到对应边界并判故障 / segment 4, the infinite gate by the self difference
IF (fIn - fIn) <> (fIn - fIn) THEN // 无穷处 fIn − fIn 产 NaN，有限值恒为零 / an infinite input yields NaN from the self difference while a finite one yields zero
    bNonFinite := TRUE; // 置非有限标志 / raise the non finite flag
    bClamped := TRUE; // 钳边界已生效 / the boundary clamp took effect
    bValid := FALSE; // 结果不可用（三件套之一，R258）/ the result is not usable
    IF fIn > DL_R2I_ZERO THEN // 正无穷 / the positive infinity
        nOut := nHi; // 钳上界 [−] / clamp to the ceiling
    ELSE // 负无穷 / the negative infinity
        nOut := nLo; // 钳下界 [−] / clamp to the floor
    END_IF
    eErr := 16#0001_064F; // 故障级：输入非有限 / fault grade, the input is not finite
    bError := TRUE; // 同拍置故障标志（R45 配对）/ raise the fault flag on the same scan
    RETURN; // 早退 / early return
END_IF

// 段 5｜判据④⑤先钳后转：转换前必须落域内（边界二，R151）/ segment 5, clamp before the conversion
fLo := INT_TO_LREAL(nLo); // 下界实数形式 [−] / the floor in real form
fHi := INT_TO_LREAL(nHi); // 上界实数形式 [−] / the ceiling in real form
IF fIn < fLo THEN // 越下界 / below the floor
    nOut := nLo; // 钳下界 [−] / clamp to the floor
    bClamped := TRUE; // 置钳位标志 / raise the clamp flag
    eErr := 16#0001_064E; // 信息级：越下界已钳位 / informational, below the floor and clamped
ELSIF fIn > fHi THEN // 越上界 / above the ceiling
    nOut := nHi; // 钳上界 [−] / clamp to the ceiling
    bClamped := TRUE; // 置钳位标志 / raise the clamp flag
    eErr := 16#0001_064E; // 信息级：越上界已钳位 / informational, above the ceiling and clamped
ELSE // 域内：向零截断（四舍五入口径归 FC_DL_RoundSat）/ inside the domain, truncate toward zero
    nOut := LREAL_TO_INT(fIn); // 向零截断（-0.5 → 0，非 -1）[−] / truncated toward zero, minus a half gives zero
END_IF

// 段 6｜统一出口（信息级钳位不置 bError，R285）/ segment 6, the unified outlet without a fault flag
bValid := TRUE; // 域内或钳位输出均可用 / an in-domain or clamped output is usable
FC_DL_RealToIntSat := TRUE; // 返回成功 / return success
END_FUNCTION

(* ---- FC_DL_RealToLintSat.st ---- *)
(*
    FC_DL_RealToLintSat —— REAL 到 LINT 域外饱和转换
    ------------------------------------------------------------------
    分类      : DL_MathData / Convert
    前缀      : FC_DL_
    版本      : 1.0.0
    溯源      : IEC 61131-3 标准语义的道莅防御性实现
                （接口语义由 IEC 61131-3 定义，内部委托平台内建 REAL_TO_LREAL、TRUNC 与 LREAL_TO_LINT，
                  外围统一错误码 / 钳位 / 双语文档；clean-room 重写，
                  未复制任何闭源厂商源码，参考实现仅限 MIT/Apache 许可）
    平台      : 纯 IEC 61131-3，CODESYS / TwinCAT / InoProShop 通用
    作者      : 道莅代码库 · PLC编程专家（R17）
    ------------------------------------------------------------------
    功能说明  : 将 REAL 防御性转换为 LINT 并作为返回值输出；
                非有限输入（NaN 或 ±INF）判为故障级 16#0001_02F1，返回 0 且 bValid=FALSE；
                取整取向声明：向零截断（TRUNC 语义）后钳位，与 R16 FC_DL_LrealToDintSat 同口径；
                升位先行：先 REAL_TO_LREAL 升位再与 LREAL 域界比较，
                禁用 REAL 常量直接比较（REAL 尾数仅 24 位，域界值本身不可精确表示，会漏判）；
                域外按方向饱和（上界 9223372036854775807 / 下界负向极值）
                并置信息级 16#0001_022E；下界用 -DL_LINT_MAX - 1 计算式，禁负数字面量直写；
                钳位方向：双侧饱和，绝不回绕。
    错误码    : 16#0001_022E 输入超 LINT 域，已按符号饱和——信息级，正常防御
                16#0001_022F 预留禁用（信息级，不得挪用）
                16#0001_02F1 非有限输入（NaN 或 ±INF）——故障级，返回 0
                16#0001_02F2 预留禁用（故障级，不得挪用）
                16#0001_02F3 预留禁用（故障级，不得挪用）
    状态机    : R6 标注 N/A —— 本组件为纯函数无顺序状态机，无 CASE 可写，非法状态不可能出现，故以本节说明替代 ELSE 兜底
    修订记录  : 2026-11-16 v1.0.0 首次入库（R17）
*)
FUNCTION FC_DL_RealToLintSat : LINT
VAR_INPUT
    fIn : REAL; // 待转换浮点值，建议域 ±9.2E18（非有限拦截，域外饱和） [无量纲] / floating value to convert, suggested domain +/-9.2E18 [dimensionless]
END_VAR
VAR_OUTPUT
    eErr   : UDINT; // 错误码，0=正常 / error id, 0=ok
    bError : BOOL;  // 是否出错，eErr 非 0 时为 TRUE / error flag, TRUE when eErr is nonzero
    bValid : BOOL;  // 输出是否有效可用 / output valid flag
END_VAR
VAR CONSTANT
    DL_LINT_MAX_LR : LREAL := 9.2233720368547758E18;  // LINT 域上界在 LREAL 域的精确可表近似值 [无量纲] / LINT upper bound represented in LREAL [dimensionless]
    DL_LINT_MAX    : LINT  := 9223372036854775807;    // LINT 上界饱和输出值 [无量纲] / LINT upper saturation output [dimensionless]
    DL_LINT_ZERO   : LINT  := 0;                      // 故障缺省返回值 [无量纲] / fault default return value [dimensionless]
    DL_REAL_INF_GUARD : LREAL := 4.0E38;              // REAL 域 ±INF 判定阈值，高于 REAL 最大有限值 3.402823E38 [无量纲] / REAL +/-INF guard above max finite REAL
END_VAR
VAR
    fLr        : LREAL; // 升位后的 LREAL 中间量 [无量纲] / widened LREAL intermediate [dimensionless]
    bNonFinite : BOOL;  // 非有限（NaN 或 ±INF）判定结果 / non-finite (NaN or +/-INF) detection result
END_VAR

// 段 1｜返回值与错误状态预置 / segment 1, preset return value and error status
FC_DL_RealToLintSat := DL_LINT_ZERO; // 故障缺省返回 0 [无量纲] / fault default 0 [dimensionless]
eErr   := 0;     // 预置无错误 / preset no error
bError := FALSE; // 预置无故障 / preset no fault
bValid := FALSE; // 预置输出无效，通过三路闸后置位 / preset invalid, set TRUE after the three gates

// 段 2｜非有限防御闸 / segment 2, non-finite guard
bNonFinite := (fIn <> fIn) OR (fIn > DL_REAL_INF_GUARD) OR (fIn < -DL_REAL_INF_GUARD); // 非有限判定（NaN 自不等 + 安全幅值判 ±INF） [无量纲] / non-finite check (NaN by self-inequality, +/-INF by safe magnitude) [dimensionless]
IF bNonFinite THEN
    eErr := 16#0001_02F1; // 非有限输入故障码 / non-finite input fault id
    bError := TRUE;       // 置故障标志 / raise error flag
    bValid := FALSE;      // 输出不可用 / output not usable
    RETURN;               // 故障级提前返回，保持缺省 0 / early return on fault, keep default 0
END_IF

// 段 3｜升位与域外判定饱和 / segment 3, widening and out-of-domain saturation
fLr := REAL_TO_LREAL(fIn); // 升位先行，REAL 域界值本身不可精确表示，直接用 REAL 比较会漏判 [无量纲] / widen first, REAL cannot represent the bound exactly so comparing in REAL would miss the overflow [dimensionless]
IF fLr > DL_LINT_MAX_LR THEN
    FC_DL_RealToLintSat := DL_LINT_MAX; // 上界饱和至 LINT 上界 [无量纲] / saturate to the LINT upper bound [dimensionless]
    eErr := 16#0001_022E;               // 信息级：域外饱和，正常防御 / info level: out-of-domain saturation, normal defence
    bError := FALSE;                    // 信息级不置故障 / info level never raises fault
    bValid := TRUE;                     // 饱和值本身有效可用 / the saturated value itself is valid
    RETURN;                             // 饱和即出口 / saturation is the exit
END_IF
IF fLr < -DL_LINT_MAX_LR THEN
    FC_DL_RealToLintSat := -DL_LINT_MAX - 1; // 下界饱和，用计算式书写，等于 LINT 最小值 [无量纲] / saturate to the LINT minimum, written as a computed expression [dimensionless]
    eErr := 16#0001_022E;                    // 上下共用同一业务语义码，方向写进头注释 / both directions share one business-semantics code, directions documented in the header
    bError := FALSE;                         // 信息级不置故障 / info level never raises fault
    bValid := TRUE;                          // 饱和值本身有效可用 / the saturated value itself is valid
    RETURN;                                  // 饱和即出口 / saturation is the exit
END_IF

// 段 4｜域内向零截断与委托转换（末段） / segment 4, in-domain truncate-toward-zero and delegated conversion (final)
FC_DL_RealToLintSat := LREAL_TO_LINT(TRUNC(fLr)); // 先 TRUNC 成整值 LREAL 再转，取向恒为向零截断，规避内建舍入取向差异 [无量纲] / TRUNC to an integral LREAL before converting, always truncates toward zero and avoids built-in rounding differences [dimensionless]
eErr   := 0;     // 域内无错误 / in-domain, no error
bError := FALSE; // 信息级不置故障 / info level never raises fault
bValid := TRUE;  // 域内输出有效可用 / in-domain output is valid
END_FUNCTION

(* ---- FC_DL_RealToRealSat.st ---- *)
(*
    FC_DL_RealToRealSat —— LREAL 到 REAL 饱和防御降型
    ------------------------------------------------------------------
    分类      : DL_MathData / Convert
    前缀      : FC_DL_
    版本      : 1.0.0
    溯源      : IEC 61131-3 标准语义的道莅防御性实现
                （内部委托平台内建 LREAL_TO_REAL 转换语义，外围统一错误码/钳位/
                  双语文档；未复制任何闭源厂商源码，参考实现仅限 MIT/Apache 许可）
    平台      : 纯 IEC 61131-3，CODESYS / TwinCAT / InoProShop 通用
    作者      : 道莅代码库 · PLC编程专家（R40）
    ------------------------------------------------------------------
    功能说明  : 将 LREAL 输入防御性降型为 REAL 并作为返回值输出，转换内核
                委托平台内建 LREAL_TO_REAL，不重实现任何转换内核；
                非有限输入（NaN 或 ±Inf）判为故障级 16#0001_03CE，返回 0.0 且
                bValid=FALSE（非有限值参与降型在三平台行为不一致，一律拦截）；
                幅值越 REAL 域钳位：|fIn| 大于 REAL 最大有限值
                3.4028234663852886E38 时钳至 ±REAL 最大有限值，置信息级 16#0001_0495；
                判定阈值取 REAL 最大有限值的 LREAL 精度字面量（可表且不低于真值），
                阈值等于真上界，不存在近似假阳性带（R15 口径自证）；
                转换前置域闸（先判域后转换）：域闸命中不调内建转换，
                保证 LREAL_TO_REAL 只接收域内可表值，杜绝降型产出 Inf；
                信息级码属正常防御：bError=FALSE、bValid=TRUE，输出钳位后防御值。
    错误码    : 16#0001_03CE 非有限输入（NaN 或 ±Inf）或域闸后的转换复检失败——故障级，返回 0.0
                16#0001_0495 输入幅值超 REAL 最大有限值，已钳至 ±3.4028234663852886E38——信息级，正常防御
                （R90 反证句：幅值钳位场景无法由故障级组合观测——钳位输出 bValid=TRUE 且
                  值为有限边界值，与域内转换的输出组合（bValid=TRUE）在幅值贴近 REAL 上界时
                  仅凭返回值无法区分「原值近似」与「已钳位」，故占信息码）
    非有限口径 : NaN 用自不等 f <> f，±Inf 用 (f − f) <> (f − f) 差值自减判定（R15）。
    状态机    : R6 标注 N/A —— 本组件为纯函数无顺序状态机，无 CASE 可写，
                非法状态不可能出现，故以本节说明替代 ELSE 兜底
    修订记录  : 2026-11-19 v1.0.0 首次入库（R40 · 批 2 · T0 快车道）
*)
FUNCTION FC_DL_RealToRealSat : REAL
VAR_INPUT
    fIn : LREAL; // 待降型输入 [无量纲] ｜ input to down-convert
END_VAR
VAR_OUTPUT
    eErr   : UDINT; // 错误码，0=正常，16#0001_04XX=信息级，16#0001_03XX=故障级 ｜ error id, 0=ok, 16#0001_04XX=info, 16#0001_03XX=fault
    bError : BOOL;  // 是否出错，eErr 落故障级时为 TRUE ｜ fault flag, TRUE when eErr is fault level
    bValid : BOOL;  // 输出是否有效可用 ｜ output valid flag
END_VAR
VAR CONSTANT
    DL_REAL_MAX_FIN : LREAL := 3.4028234663852886E38; // REAL 最大有限值（LREAL 精度字面量，恰为真上界）[无量纲] ｜ largest finite REAL as an LREAL literal (the true upper bound)
END_VAR
VAR
    bNonFinite : BOOL; // 非有限（NaN 或 ±Inf）判定结果 ｜ non-finite (NaN or +/-Inf) detection result
    fOut       : REAL; // 降型结果暂存，供出口复检 ｜ staging of the converted result for exit recheck
END_VAR

// 段 1｜返回值与错误状态预置 ｜ segment 1, preset return value and error status
FC_DL_RealToRealSat := 0.0; // 故障缺省返回 0 [无量纲] ｜ fault default returns 0
eErr   := 0;     // 预置无错误 ｜ preset no error
bError := FALSE; // 预置无故障 ｜ preset no fault
bValid := FALSE; // 预置无效，通过防御闸后置位 ｜ preset invalid, set TRUE after guard passes
fOut   := 0.0;   // 暂存清零 ｜ clear the staging value

// 段 2｜非有限防御闸（命中不调内建转换，早退） ｜ segment 2, non-finite guard (early return, no built-in conversion)
bNonFinite := (fIn <> fIn) OR ((fIn - fIn) <> (fIn - fIn)); // NaN 自不等 + 差值自减判 ±Inf [无量纲] ｜ NaN by self-inequality, +/-Inf by self-subtraction
IF bNonFinite THEN
    FC_DL_RealToRealSat := 0.0; // 故障级返回 0 [无量纲] ｜ fault level returns 0
    eErr   := 16#0001_03CE;     // 非有限输入故障码 ｜ non-finite input fault id
    bError := TRUE;             // 置故障标志（R45 配对）｜ raise the fault flag (R45 pairing)
    bValid := FALSE;            // 输出无效 ｜ output invalid
    RETURN;                     // 早退，不调内建转换 ｜ early return, no built-in conversion
END_IF

// 段 3｜幅值域闸与降型转换（先判域后转换） ｜ segment 3, magnitude domain gate and down-conversion (domain check before conversion)
IF fIn > DL_REAL_MAX_FIN THEN
    fOut := 3.4028235E38;     // 正幅值越域钳至 REAL 最大有限值 [无量纲] ｜ positive magnitude clamped to the largest finite REAL
    eErr := 16#0001_0495;     // 信息级：幅值越 REAL 域已钳位 ｜ info level: magnitude beyond the REAL domain, clamped
ELSIF fIn < -DL_REAL_MAX_FIN THEN
    fOut := -3.4028235E38;    // 负幅值越域钳至 REAL 最小有限值 [无量纲] ｜ negative magnitude clamped to the smallest finite REAL
    eErr := 16#0001_0495;     // 信息级：幅值越 REAL 域已钳位（双侧共用幅值钳位码，方向由输出符号还原）｜ info level: clamped (both sides share the magnitude code, direction recovered from the output sign)
ELSE
    fOut := LREAL_TO_REAL(fIn); // 域内委托平台内建降型转换 ｜ in-domain delegate to the built-in down-conversion
    eErr := 0;                  // 域内无错误 ｜ in-domain, no error
END_IF

// 段 4｜结果复检兜底（理论不可达：域闸后的降型恒产出有限 REAL） ｜ segment 4, exit recheck (unreachable: in-domain down-conversion always yields a finite REAL)
IF (fOut <> fOut) OR ((LREAL_TO_REAL(fOut) - LREAL_TO_REAL(fOut)) <> (LREAL_TO_REAL(fOut) - LREAL_TO_REAL(fOut))) THEN
    FC_DL_RealToRealSat := 0.0; // 复检失败按非有限处置 [无量纲] ｜ recheck failure treated as non-finite
    eErr   := 16#0001_03CE;     // 复用非有限码（同因同码，不新占码位）｜ reuse the non-finite code (same cause, no new code)
    bError := TRUE;             // 置故障标志 ｜ raise the fault flag
    bValid := FALSE;            // 输出无效 ｜ output invalid
    RETURN;                     // 早退 ｜ early return
END_IF

// 段 5｜出口装配 ｜ segment 5, exit assembly
FC_DL_RealToRealSat := fOut; // 降型结果直通 ｜ converted result pass-through
bError := FALSE;             // 信息级钳位不置故障，故障分支已提前返回 ｜ info-level clamp never raises fault, fault branch has returned
bValid := TRUE;              // 域内或钳位输出均有效可用 ｜ in-domain or clamped output is valid
END_FUNCTION

(* ---- FC_DL_RealToUdintSat.st ---- *)
(*
    FC_DL_RealToUdintSat —— REAL 到 UDINT 饱和防御转换
    ------------------------------------------------------------------
    分类      : DL_MathData / Convert
    前缀      : FC_DL_
    版本      : 1.0.0
    溯源      : IEC 61131-3 标准语义的道莅防御性实现
                （内部委托平台内建函数，外围统一错误码/钳位/双语文档；
                  未复制任何闭源厂商源码，参考实现仅限 MIT/Apache 许可）
    平台      : 纯 IEC 61131-3，CODESYS / TwinCAT / InoProShop 通用
    作者      : 道莅代码库 · PLC编程专家（R16）
    ------------------------------------------------------------------
    功能说明  : 将 REAL 输入防御性转换为 UDINT 并作为返回值输出；
                非有限输入（NaN 或 ±INF）判为故障级 16#0001_0294，返回 0 且 bValid=FALSE；
                fIn < 0 时钳位至 0，置信息级 16#0001_01C4（UDINT 无符号，负值不可表）；
                fIn 超出 UDINT 上界 4294967295 时钳位至上界，置信息级 16#0001_01C5；
                钳位方向：下界 0 / 上界 4294967295（双侧饱和）；
                ±INF 采用平台安全幅值比较判定（阈值高于 REAL 最大有限值 3.402823E38），NaN 用 fIn <> fIn 自不等判定；
                域内转换委托平台内建 REAL_TO_UDINT 语义，不重实现数学内核；
                信息级码属正常防御：bError=FALSE、bValid=TRUE，输出钳位后防御值。
    错误码    : 16#0001_0294 非有限输入（NaN 或 ±INF）——故障级，返回 0
                16#0001_01C4 负值输入，已钳位至 0——信息级，正常防御
                16#0001_01C5 输入超 UDINT 上界，已钳位至 4294967295——信息级，正常防御
                16#0001_0295 预留禁用（故障级，不得挪用）
                16#0001_0296 预留禁用（故障级，不得挪用）
    状态机    : R6 标注 N/A —— 本组件为纯函数无顺序状态机，无 CASE 可写，非法状态不可能出现，故以本节说明替代 ELSE 兜底
    修订记录  : 2026-11-16 v1.0.0 首次入库（R16）
*)
FUNCTION FC_DL_RealToUdintSat : UDINT
VAR_INPUT
    fIn : REAL; // 待转换输入 [无量纲] / input value to convert
END_VAR
VAR_OUTPUT
    eErr   : UDINT; // 错误码，0=正常 / error id, 0=ok
    bError : BOOL;  // 是否出错，eErr 非 0 时为 TRUE / error flag, TRUE when eErr is nonzero
    bValid : BOOL;  // 输出是否有效可用 / output valid flag
END_VAR
VAR CONSTANT
    DL_UDINT_MAX      : LREAL := 4.294967295E9; // UDINT 域上界 4294967295，LREAL 承载 [无量纲] / UDINT upper bound 4294967295 carried in LREAL
    DL_REAL_INF_GUARD : LREAL := 4.0E38;        // REAL 域 ±INF 判定阈值，高于 REAL 最大有限值 3.402823E38 [无量纲] / REAL +/-INF guard above max finite REAL 3.402823E38
END_VAR
VAR
    bNonFinite : BOOL; // 非有限（NaN 或 ±INF）判定结果 / non-finite (NaN or +/-INF) detection result
END_VAR

// 段 1｜返回值与错误状态预置 / segment 1, preset return value and error status
FC_DL_RealToUdintSat := 0; // 故障缺省返回 0 [无量纲] / fault default returns 0
eErr   := 0;     // 预置无错误 / preset no error
bError := FALSE; // 预置无故障 / preset no fault
bValid := FALSE; // 预置无效，通过防御闸后置位 / preset invalid, set TRUE after guard passes

// 段 2｜非有限防御闸 / segment 2, non-finite guard
bNonFinite := (fIn <> fIn) OR (fIn > DL_REAL_INF_GUARD) OR (fIn < -DL_REAL_INF_GUARD); // NaN 自不等判定，±INF 用安全幅值比较 [无量纲] / NaN by self-inequality, +/-INF by safe magnitude compare
IF bNonFinite THEN
    FC_DL_RealToUdintSat := 0; // 故障级返回 0 [无量纲] / fault level returns 0
    eErr   := 16#0001_0294;    // 非有限输入故障码 / non-finite input fault id
    bError := TRUE;            // 置故障标志 / set fault flag
    bValid := FALSE;           // 输出无效 / output invalid
    RETURN;                    // 立即返回 / immediate return
END_IF

// 段 3｜双侧饱和钳位与主体转换（末段） / segment 3, double-side saturating clamp and main conversion (final)
IF fIn < 0.0 THEN
    FC_DL_RealToUdintSat := 0;      // 负值钳位至 0（UDINT 无符号语义） / negative input clamped to 0 (UDINT is unsigned)
    eErr := 16#0001_01C4;           // 信息级：负值已钳零 / info level: negative input clamped to zero
ELSIF fIn > DL_UDINT_MAX THEN
    FC_DL_RealToUdintSat := 16#FFFFFFFF; // 正向钳位至 UDINT 上界 4294967295 / clamp to UDINT upper bound 4294967295
    eErr := 16#0001_01C5;                // 信息级：超上界已钳位 / info level: above upper bound, clamped
ELSE
    FC_DL_RealToUdintSat := REAL_TO_UDINT(fIn); // 域内委托平台内建 _TO_ 转换语义 / in-domain delegate to built-in _TO_ conversion
    eErr := 0; // 域内无错误 / in-domain, no error
END_IF
bError := FALSE; // 信息级钳位不置故障，故障分支已提前返回 / info-level clamp never raises fault, fault branch has returned
bValid := TRUE;  // 域内或钳位输出均有效可用 / in-domain or clamped output is valid
END_FUNCTION
